           "Control_DB"."Carrousel_Order Table".Task_Data_Available := TRUE;//#System.OrderTable[#Roller_To_Roller_CurrentOrder].OPC_Control.Task_Data_Available; // Send the Task Data Available from WCS 
           "Control_DB"."Carrousel_Order Table".Task_Type := #System.OrderTable[#RTR_P1P2_CurrentOrder].OPC_Control.Task_Type; //  Send the Task Type - Roller to Roller Conveyor = Task Type = 6
           "Control_DB"."Carrousel_Order Table".Task_ID := #System.OrderTable[#RTR_P1P2_CurrentOrder].OPC_Control.Task_ID; // Send the Task ID number;
           "Control_DB"."Carrousel_Order Table".Task_Metadata := #System.OrderTable[#RTR_P1P2_CurrentOrder].OPC_Control.Task_Metadata; // Send the Task Metadata Unique identifier
           "Control_DB"."Carrousel_Order Table".Source_Location := #System.OrderTable[#RTR_P1P2_CurrentOrder].OPC_Control.Source_Location; // Send the Source Location from the Conveyor
           "Control_DB"."Carrousel_Order Table".Destination_Location := #System.OrderTable[#RTR_P1P2_CurrentOrder].OPC_Control.Destination_Location; // Send the Destination Location to the Conveyor;
           #RTR_P1P2_WatchdogStart := true;


       END_IF;

       //RUNNING
       IF (#Cnv_PopUp_1.Running OR #Cnv_PopUp_2.Running) AND #System.Auto_Man THEN
           #System.OrderTable[#RTR_P1P2_CurrentOrder].Status := #RUNNING_STATUS;
       END_IF;

       //Cancel order
       IF #Canceling AND NOT (#Cnv_PopUp_1.Running OR #Cnv_PopUp_2.Running) AND #RTR_P1P2_CurrentOrder <> 0
       THEN
           #System.OrderTable[#RTR_P1P2_CurrentOrder].Status := #CANCELED_STATUS;
           #System.OrderTable[#RTR_P1P2_CurrentOrder].CompleteTime := #CurrentTime;
           #RTR_P1P2_CurrentOrder := 0;

           "Control_DB"."Profiling Station".Start := FALSE;

           "Control_DB"."Carrousel_Order Table".Task_Data_Available := FALSE; // Send the Task Data Available from WCS 
           "Control_DB"."Carrousel_Order Table".Task_Type := 0; //  Send the Task Type - Roller to Roller Conveyor = Task Type = 6
           "Control_DB"."Carrousel_Order Table".Task_ID := 0; // Send the Task ID number;
           "Control_DB"."Carrousel_Order Table".Task_Metadata := ''; // Send the Task Metadata Unique identifier
           "Control_DB"."Carrousel_Order Table".Source_Location := 0; // Send the Source Location from the Conveyor
           "Control_DB"."Carrousel_Order Table".Destination_Location := 0; // Send the Destination Location to the Conveyor;

       END_IF;

       //Error
       IF (#Cnv_PopUp_1.Error OR #Cnv_PopUp_2.Error) THEN
           //#Cnv_Entry.Instruction.Execute := FALSE;
           "Control_DB"."Profiling Station".Start := FALSE;

           "Control_DB"."Carrousel_Order Table".Task_Data_Available := FALSE; // Send the Task Data Available from WCS 
           "Control_DB"."Carrousel_Order Table".Task_Type := 0; //  Send the Task Type - Roller to Roller Conveyor = Task Type = 6
           "Control_DB"."Carrousel_Order Table".Task_ID := 0; // Send the Task ID number;
           "Control_DB"."Carrousel_Order Table".Task_Metadata := ''; // Send the Task Metadata Unique identifier
           "Control_DB"."Carrousel_Order Table".Source_Location := 0; // Send the Source Location from the Conveyor
           "Control_DB"."Carrousel_Order Table".Destination_Location := 0; // Send the Destination Location to the Conveyor;
           #System.OrderTable[#RTR_P1P2_CurrentOrder].ErrorID := (#Cnv_PopUp_1.Cnv_Errors.Error_Word_1
           OR #Cnv_PopUp_2.Cnv_Errors.Error_Word_1)
       ;

       END_IF;

       //MOVEMENT FINALIZED
       #RTR_P1P2DoneRTrig(CLK := "Control_DB".Movement_Completed.RTR_P1TP2);
       IF #RTR_P1P2DoneRTrig.Q THEN
           "Control_DB".Movement_Completed.RTR_P1TP2 := FALSE;
           "Control_DB"."Profiling Station".Start := FALSE;

           "Control_DB"."Carrousel_Order Table".Task_Data_Available := FALSE; // Send the Task Data Available from WCS 
           "Control_DB"."Carrousel_Order Table".Task_Type := 0; //  Send the Task Type - Roller to Roller Conveyor = Task Type = 6
           "Control_DB"."Carrousel_Order Table".Task_ID := 0; // Send the Task ID number;
           "Control_DB"."Carrousel_Order Table".Task_Metadata := ''; // Send the Task Metadata Unique identifier
           "Control_DB"."Carrousel_Order Table".Source_Location := 0; // Send the Source Location from the Conveyor
           "Control_DB"."Carrousel_Order Table".Destination_Location := 0; // Send the Destination Location to the Conveyor;

           #RTR_P1P2_WatchdogStart := FALSE;
           #System.OrderTable[#RTR_P1P2_CurrentOrder].Status := #COMPLETED_STATUS;
           #System.OrderTable[#RTR_P1P2_CurrentOrder].CompleteTime := #CurrentTime;
           #RTR_P1P2_CurrentOrder := 0;
       END_IF;
   END_REGION

   REGION Roller TO Roller - Carousel Conveyors - PP3 PP4
       //Roller conveyors
       IF #System.OrderTable[1].StepNo <> 0
           AND #System.OrderTable[1].Device = #RTR_P3_TO_P4
           AND #System.OrderTable[1].Status = #QUEUED_STATUS
           AND NOT (#Cnv_PopUp_3.Running OR #Cnv_PopUp_4.Running)
           AND NOT #System.Error
           AND NOT #Canceling

       THEN
           #RTR_P3P4_CurrentOrder := 1;
       END_IF;
       IF #System.OrderTable[#RTR_P3P4_CurrentOrder].StepNo <> 0
           AND #System.OrderTable[#RTR_P3P4_CurrentOrder].Device = #RTR_P3_TO_P4
           AND #System.OrderTable[#RTR_P3P4_CurrentOrder].Status = #QUEUED_STATUS
           AND NOT (#Cnv_PopUp_3.Running OR #Cnv_PopUp_4.Running)
           AND NOT #System.Error
           AND NOT #Canceling

       THEN
           //OPC Commands to Move Pallets - Carousel Conveyors
           // WCS => Order Table => OPC Ua Control Table


           "Control_DB"."Carrousel_Order Table".Task_Data_Available := TRUE;//#System.OrderTable[#Roller_To_Roller_CurrentOrder].OPC_Control.Task_Data_Available; // Send the Task Data Available from WCS 
           "Control_DB"."Carrousel_Order Table".Task_Type := #System.OrderTable[#RTR_P3P4_CurrentOrder].OPC_Control.Task_Type; //  Send the Task Type - Roller to Roller Conveyor = Task Type = 6
           "Control_DB"."Carrousel_Order Table".Task_ID := #System.OrderTable[#RTR_P3P4_CurrentOrder].OPC_Control.Task_ID; // Send the Task ID number;
           "Control_DB"."Carrousel_Order Table".Task_Metadata := #System.OrderTable[#RTR_P3P4_CurrentOrder].OPC_Control.Task_Metadata; // Send the Task Metadata Unique identifier
           "Control_DB"."Carrousel_Order Table".Source_Location := #System.OrderTable[#RTR_P3P4_CurrentOrder].OPC_Control.Source_Location; // Send the Source Location from the Conveyor
           "Control_DB"."Carrousel_Order Table".Destination_Location := #System.OrderTable[#RTR_P3P4_CurrentOrder].OPC_Control.Destination_Location; // Send the Destination Location to the Conveyor;
           #RTR_P3P4_WatchdogStart := true;


       END_IF;

       //RUNNING
       IF (#Cnv_PopUp_4.Running OR #Cnv_PopUp_3.Running) AND #System.Auto_Man THEN
           #System.OrderTable[#RTR_P3P4_CurrentOrder].Status := #RUNNING_STATUS;
       END_IF;

       //Cancel order
       IF #Canceling AND NOT (#Cnv_PopUp_4.Running OR #Cnv_PopUp_3.Running) AND #RTR_P3P4_CurrentOrder <> 0
       THEN
           #System.OrderTable[#RTR_P3P4_CurrentOrder].Status := #CANCELED_STATUS;
           #System.OrderTable[#RTR_P3P4_CurrentOrder].CompleteTime := #CurrentTime;
           #RTR_P3P4_CurrentOrder := 0;


           "Control_DB"."Carrousel_Order Table".Task_Data_Available := FALSE; // Send the Task Data Available from WCS 
           "Control_DB"."Carrousel_Order Table".Task_Type := 0; //  Send the Task Type - Roller to Roller Conveyor = Task Type = 6
           "Control_DB"."Carrousel_Order Table".Task_ID := 0; // Send the Task ID number;
           "Control_DB"."Carrousel_Order Table".Task_Metadata := ''; // Send the Task Metadata Unique identifier
           "Control_DB"."Carrousel_Order Table".Source_Location := 0; // Send the Source Location from the Conveyor
           "Control_DB"."Carrousel_Order Table".Destination_Location := 0; // Send the Destination Location to the Conveyor;

       END_IF;

       //Error
       IF (#Cnv_PopUp_4.Error OR #Cnv_PopUp_3.Error) THEN
           //#Cnv_Entry.Instruction.Execute := FALSE;

           "Control_DB"."Carrousel_Order Table".Task_Data_Available := FALSE; // Send the Task Data Available from WCS 
           "Control_DB"."Carrousel_Order Table".Task_Type := 0; //  Send the Task Type - Roller to Roller Conveyor = Task Type = 6
           "Control_DB"."Carrousel_Order Table".Task_ID := 0; // Send the Task ID number;
           "Control_DB"."Carrousel_Order Table".Task_Metadata := ''; // Send the Task Metadata Unique identifier
           "Control_DB"."Carrousel_Order Table".Source_Location := 0; // Send the Source Location from the Conveyor
           "Control_DB"."Carrousel_Order Table".Destination_Location := 0; // Send the Destination Location to the Conveyor;
           #System.OrderTable[#RTR_P3P4_CurrentOrder].ErrorID := (#Cnv_PopUp_3.Cnv_Errors.Error_Word_1
           OR #Cnv_PopUp_4.Cnv_Errors.Error_Word_1)
           ;

       END_IF;

       //MOVEMENT FINALIZED
       #RTR_P3P4DoneRTrig(CLK := "Control_DB".Movement_Completed.RTR_P3TP4);
       IF #RTR_P3P4DoneRTrig.Q THEN
           "Control_DB".Movement_Completed.RTR_P3TP4 := FALSE;

           "Control_DB"."Carrousel_Order Table".Task_Data_Available := FALSE; // Send the Task Data Available from WCS 
           "Control_DB"."Carrousel_Order Table".Task_Type := 0; //  Send the Task Type - Roller to Roller Conveyor = Task Type = 6
           "Control_DB"."Carrousel_Order Table".Task_ID := 0; // Send the Task ID number;
           "Control_DB"."Carrousel_Order Table".Task_Metadata := ''; // Send the Task Metadata Unique identifier
           "Control_DB"."Carrousel_Order Table".Source_Location := 0; // Send the Source Location from the Conveyor
           "Control_DB"."Carrousel_Order Table".Destination_Location := 0; // Send the Destination Location to the Conveyor;

           #RTR_P3P4_WatchdogStart := FALSE;
           #System.OrderTable[#RTR_P3P4_CurrentOrder].Status := #COMPLETED_STATUS;
           #System.OrderTable[#RTR_P3P4_CurrentOrder].CompleteTime := #CurrentTime;
           #RTR_P3P4_CurrentOrder := 0;
       END_IF;
   END_REGION

   REGION Roller TO Roller - Carousel Conveyors - PP4 to outbound
       //Roller conveyors
       IF #System.OrderTable[1].StepNo <> 0
           AND #System.OrderTable[1].Device = #RTR_P4TO
           AND #System.OrderTable[1].Status = #QUEUED_STATUS
           AND NOT (#Cnv_PopUp_4.Running OR #Cnv_Exit.Running)
           AND NOT #System.Error
           AND NOT #Canceling

       THEN
           #RTR_P4TO_CurrentOrder := 1;
       END_IF;
       IF #System.OrderTable[#RTR_P4TO_CurrentOrder].StepNo <> 0
           AND #System.OrderTable[#RTR_P4TO_CurrentOrder].Device = #RTR_P4TO
           AND #System.OrderTable[#RTR_P4TO_CurrentOrder].Status = #QUEUED_STATUS
           AND NOT (#Cnv_PopUp_4.Running OR #Cnv_Exit.Running)
           AND NOT #System.Error
           AND NOT #Canceling

       THEN
           //OPC Commands to Move Pallets - Carousel Conveyors
           // WCS => Order Table => OPC Ua Control Table


           "Control_DB"."Carrousel_Order Table".Task_Data_Available := TRUE;//#System.OrderTable[#Roller_To_Roller_CurrentOrder].OPC_Control.Task_Data_Available; // Send the Task Data Available from WCS 
           "Control_DB"."Carrousel_Order Table".Task_Type := #System.OrderTable[#RTR_P4TO_CurrentOrder].OPC_Control.Task_Type; //  Send the Task Type - Roller to Roller Conveyor = Task Type = 6
           "Control_DB"."Carrousel_Order Table".Task_ID := #System.OrderTable[#RTR_P4TO_CurrentOrder].OPC_Control.Task_ID; // Send the Task ID number;
           "Control_DB"."Carrousel_Order Table".Task_Metadata := #System.OrderTable[#RTR_P4TO_CurrentOrder].OPC_Control.Task_Metadata; // Send the Task Metadata Unique identifier
           "Control_DB"."Carrousel_Order Table".Source_Location := #System.OrderTable[#RTR_P4TO_CurrentOrder].OPC_Control.Source_Location; // Send the Source Location from the Conveyor
           "Control_DB"."Carrousel_Order Table".Destination_Location := #System.OrderTable[#RTR_P4TO_CurrentOrder].OPC_Control.Destination_Location; // Send the Destination Location to the Conveyor;
           #RTR_P4TO_WatchdogStart := true;


       END_IF;

       //RUNNING
       IF (#Cnv_PopUp_4.Running OR #Cnv_Exit.Running) AND #System.Auto_Man THEN
           #System.OrderTable[#RTR_P4TO_CurrentOrder].Status := #RUNNING_STATUS;
       END_IF;

       //Cancel order
       IF #Canceling AND NOT (#Cnv_PopUp_4.Running OR #Cnv_Exit.Running) AND #RTR_P4TO_CurrentOrder <> 0
       THEN
           #System.OrderTable[#RTR_P4TO_CurrentOrder].Status := #CANCELED_STATUS;
           #System.OrderTable[#RTR_P4TO_CurrentOrder].CompleteTime := #CurrentTime;
           #RTR_P4TO_CurrentOrder := 0;


           "Control_DB"."Carrousel_Order Table".Task_Data_Available := FALSE; // Send the Task Data Available from WCS 
           "Control_DB"."Carrousel_Order Table".Task_Type := 0; //  Send the Task Type - Roller to Roller Conveyor = Task Type = 6
           "Control_DB"."Carrousel_Order Table".Task_ID := 0; // Send the Task ID number;
           "Control_DB"."Carrousel_Order Table".Task_Metadata := ''; // Send the Task Metadata Unique identifier
           "Control_DB"."Carrousel_Order Table".Source_Location := 0; // Send the Source Location from the Conveyor
           "Control_DB"."Carrousel_Order Table".Destination_Location := 0; // Send the Destination Location to the Conveyor;

       END_IF;

       //Error
       IF (#Cnv_PopUp_4.Error OR #Cnv_Exit.Error) THEN
           //#Cnv_Entry.Instruction.Execute := FALSE;

           "Control_DB"."Carrousel_Order Table".Task_Data_Available := FALSE; // Send the Task Data Available from WCS 
           "Control_DB"."Carrousel_Order Table".Task_Type := 0; //  Send the Task Type - Roller to Roller Conveyor = Task Type = 6
           "Control_DB"."Carrousel_Order Table".Task_ID := 0; // Send the Task ID number;
           "Control_DB"."Carrousel_Order Table".Task_Metadata := ''; // Send the Task Metadata Unique identifier
           "Control_DB"."Carrousel_Order Table".Source_Location := 0; // Send the Source Location from the Conveyor
           "Control_DB"."Carrousel_Order Table".Destination_Location := 0; // Send the Destination Location to the Conveyor;
           #System.OrderTable[#RTR_P3P4_CurrentOrder].ErrorID := (#Cnv_PopUp_3.Cnv_Errors.Error_Word_1
           OR #Cnv_PopUp_4.Cnv_Errors.Error_Word_1)
           ;

       END_IF;

       //MOVEMENT FINALIZED
       #RTR_P4TODoneRTrig(CLK := "Control_DB".Movement_Completed.RTR_P4TO);
       IF #RTR_P4TODoneRTrig.Q THEN
           "Control_DB".Movement_Completed.RTR_P4TO := FALSE;

           "Control_DB"."Carrousel_Order Table".Task_Data_Available := FALSE; // Send the Task Data Available from WCS 
           "Control_DB"."Carrousel_Order Table".Task_Type := 0; //  Send the Task Type - Roller to Roller Conveyor = Task Type = 6
           "Control_DB"."Carrousel_Order Table".Task_ID := 0; // Send the Task ID number;
           "Control_DB"."Carrousel_Order Table".Task_Metadata := ''; // Send the Task Metadata Unique identifier
           "Control_DB"."Carrousel_Order Table".Source_Location := 0; // Send the Source Location from the Conveyor
           "Control_DB"."Carrousel_Order Table".Destination_Location := 0; // Send the Destination Location to the Conveyor;

           #RTR_P4TO_WatchdogStart := FALSE;
           #System.OrderTable[#RTR_P4TO_CurrentOrder].Status := #COMPLETED_STATUS;
           #System.OrderTable[#RTR_P4TO_CurrentOrder].CompleteTime := #CurrentTime;
           #RTR_P4TO_CurrentOrder := 0;
       END_IF;
   END_REGION




   REGION Chain to Chain - Carousel Conveyors - Pop 2 to Pop 3
       IF #System.OrderTable[1].StepNo <> 0
           AND #System.OrderTable[1].Device = #CHAIN_TO_CHAIN_DEVICE
           AND #System.OrderTable[1].Status = #QUEUED_STATUS
           AND NOT (#Cnv_PopUp_2.Running OR #Cnv_PopUp_3.Running)
           AND NOT #System.Error
           AND NOT #Canceling
           //AND #System.OrderTable[#Chain_To_Chain_CurrentOrder].Status <> #RUNNING_STATUS

       THEN
           #Chain_To_Chain_CurrentOrder := 1;
       END_IF;
       IF #System.OrderTable[#Chain_To_Chain_CurrentOrder].StepNo <> 0
           AND #System.OrderTable[#Chain_To_Chain_CurrentOrder].Device = #CHAIN_TO_CHAIN_DEVICE
           AND #System.OrderTable[#Chain_To_Chain_CurrentOrder].Status = #QUEUED_STATUS
           AND NOT (#Cnv_PopUp_2.Running OR #Cnv_PopUp_3.Running)
           AND NOT #System.Error
           AND NOT #Canceling
          // AND #System.OrderTable[#Chain_To_Chain_CurrentOrder].Status <> #RUNNING_STATUS
       THEN
           //OPC Commands to Move Pallets - Carousel Conveyors
           // WCS => Order Table => OPC Ua Control Table

           "Control_DB"."Carrousel_Order Table".Task_Data_Available := TRUE;//#System.OrderTable[#Chain_To_Chain_CurrentOrder].OPC_Control.Task_Data_Available; // Send the Task Data Available from WCS 
           "Control_DB"."Carrousel_Order Table".Task_Type := #System.OrderTable[#Chain_To_Chain_CurrentOrder].OPC_Control.Task_Type; //  Send the Task Type - Chain to Chain Conveyor = Task Type = 7
           "Control_DB"."Carrousel_Order Table".Task_ID := #System.OrderTable[#Chain_To_Chain_CurrentOrder].OPC_Control.Task_ID; // Send the Task ID number;
           "Control_DB"."Carrousel_Order Table".Task_Metadata := #System.OrderTable[#Chain_To_Chain_CurrentOrder].OPC_Control.Task_Metadata; // Send the Task Metadata Unique identifier
           "Control_DB"."Carrousel_Order Table".Source_Location := #System.OrderTable[#Chain_To_Chain_CurrentOrder].OPC_Control.Source_Location; // Send the Source Location from the Conveyor
           "Control_DB"."Carrousel_Order Table".Destination_Location := #System.OrderTable[#Chain_To_Chain_CurrentOrder].OPC_Control.Destination_Location; // Send the Destination Location to the Conveyor;
           #Chain_To_Chain_WatchdogStart := true;


       END_IF;

       //RUNNING
       IF (#Cnv_PopUp_2.Running OR #Cnv_PopUp_3.Running)AND #System.Auto_Man THEN
           //#Cnv_Entry.Instruction.Execute := FALSE;
           #System.OrderTable[#Chain_To_Chain_CurrentOrder].Status := #RUNNING_STATUS;
       END_IF;

       //Cancel order
       IF #Canceling AND NOT (#Cnv_PopUp_2.Running OR #Cnv_PopUp_3.Running) AND #Chain_To_Chain_CurrentOrder <> 0 THEN


           "Control_DB"."Carrousel_Order Table".Task_Data_Available := FALSE;//#System.OrderTable[#Chain_To_Chain_CurrentOrder].OPC_Control.Task_Data_Available; // Send the Task Data Available from WCS 
           "Control_DB"."Carrousel_Order Table".Task_Type := 0; //  Send the Task Type - Chain to Chain Conveyor = Task Type = 7
           "Control_DB"."Carrousel_Order Table".Task_ID := 0; // Send the Task ID number;
           "Control_DB"."Carrousel_Order Table".Task_Metadata := ''; // Send the Task Metadata Unique identifier
           "Control_DB"."Carrousel_Order Table".Source_Location := 0; // Send the Source Location from the Conveyor
           "Control_DB"."Carrousel_Order Table".Destination_Location := 0; // Send the Destination Location to the Conveyor;

           #System.OrderTable[#Chain_To_Chain_CurrentOrder].Status := #CANCELED_STATUS;
           #System.OrderTable[#Chain_To_Chain_CurrentOrder].CompleteTime := #CurrentTime;
           #Chain_To_Chain_CurrentOrder := 0;
           //#Cnv_Entry.Instruction.Execute := FALSE;
       END_IF;

       //Error
       IF (#Cnv_PopUp_2.Error OR #Cnv_PopUp_3.Error) THEN
           //#Cnv_Entry.Instruction.Execute := FALSE;
           //
           "Control_DB"."Carrousel_Order Table".Task_Data_Available := FALSE;//#System.OrderTable[#Chain_To_Chain_CurrentOrder].OPC_Control.Task_Data_Available; // Send the Task Data Available from WCS 
           "Control_DB"."Carrousel_Order Table".Task_Type := 0; //  Send the Task Type - Chain to Chain Conveyor = Task Type = 7
           "Control_DB"."Carrousel_Order Table".Task_ID := 0; // Send the Task ID number;
           "Control_DB"."Carrousel_Order Table".Task_Metadata := ''; // Send the Task Metadata Unique identifier
           "Control_DB"."Carrousel_Order Table".Source_Location := 0; // Send the Source Location from the Conveyor
           "Control_DB"."Carrousel_Order Table".Destination_Location := 0; // Send the Destination Location to the Conveyor;

           #System.OrderTable[#Chain_To_Chain_CurrentOrder].ErrorID := (#Cnv_PopUp_2.Cnv_Errors.Error_Word_1
                                                                        OR #Cnv_PopUp_3.Cnv_Errors.Error_Word_1);

       END_IF;

       //MOVEMENT FINALIZED
       #Chain_To_ChainDoneRTrig(CLK := "Control_DB".Movement_Completed.RTR_P2TP3);
       IF #Chain_To_ChainDoneRTrig.Q THEN
           "Control_DB".Movement_Completed.RTR_P2TP3 := FALSE;
           "Control_DB"."Carrousel_Order Table".Task_Data_Available := FALSE;//#System.OrderTable[#Chain_To_Chain_CurrentOrder].OPC_Control.Task_Data_Available; // Send the Task Data Available from WCS 
           "Control_DB"."Carrousel_Order Table".Task_Type := 0; //  Send the Task Type - Chain to Chain Conveyor = Task Type = 7
           "Control_DB"."Carrousel_Order Table".Task_ID := 0; // Send the Task ID number;
           "Control_DB"."Carrousel_Order Table".Task_Metadata := ''; // Send the Task Metadata Unique identifier
           "Control_DB"."Carrousel_Order Table".Source_Location := 0; // Send the Source Location from the Conveyor
           "Control_DB"."Carrousel_Order Table".Destination_Location := 0; // Send the Destination Location to the Conveyor;


           #Chain_To_Chain_WatchdogStart := FALSE;
           #System.OrderTable[#Chain_To_Chain_CurrentOrder].Status := #COMPLETED_STATUS;
           #System.OrderTable[#Chain_To_Chain_CurrentOrder].CompleteTime := #CurrentTime;
           #Chain_To_Chain_CurrentOrder := 0;
       END_IF;
   END_REGION

   REGION Pop4 to Pick Station - Carousel Conveyors - Pop 4 to Pick Station
       IF #System.OrderTable[1].StepNo <> 0
           AND #System.OrderTable[1].Device = #POP4_TO_PICK_DEVICE
           AND #System.OrderTable[1].Status = #QUEUED_STATUS
          // AND NOT "Control_DB".Pick_Station.Running
           AND NOT #System.Error
           AND NOT #Canceling
           AND #System.OrderTable[1].Status <> #RUNNING_STATUS
           //AND #System.OrderTable[#PickSt_To_Pop1_CurrentOrder].Status <> #RUNNING_STATUS

       THEN
           #Pop4_To_PickSt_CurrentOrder := 1;
       END_IF;
       IF #System.OrderTable[#Pop4_To_PickSt_CurrentOrder].StepNo <> 0
           AND #System.OrderTable[#Pop4_To_PickSt_CurrentOrder].Device = #POP4_TO_PICK_DEVICE
           AND #System.OrderTable[#Pop4_To_PickSt_CurrentOrder].Status = #QUEUED_STATUS
           // AND NOT "Control_DB".Pick_Station.Running
           AND NOT #System.Error
           AND NOT #Canceling
           AND #System.OrderTable[#Pop4_To_PickSt_CurrentOrder].Status <> #RUNNING_STATUS
           //AND #System.OrderTable[#PickSt_To_Pop1_CurrentOrder].Status <> #RUNNING_STATUS
       THEN
           //OPC Commands to Move Pallets - Carousel Conveyors
           // WCS => Order Table => OPC Ua Control Table

           "Control_DB"."Carrousel_Order Table".Task_Data_Available := TRUE;//#System.OrderTable[#Pop4_To_PickSt_CurrentOrder].OPC_Control.Task_Data_Available; // Send the Task Data Available from WCS 
           "Control_DB"."Carrousel_Order Table".Task_Type := #System.OrderTable[#Pop4_To_PickSt_CurrentOrder].OPC_Control.Task_Type; //  Send the Task Type - Pop4 to Pick Station Conveyor = Task Type = 8
           "Control_DB"."Carrousel_Order Table".Task_ID := #System.OrderTable[#Pop4_To_PickSt_CurrentOrder].OPC_Control.Task_ID; // Send the Task ID number;
           "Control_DB"."Carrousel_Order Table".Task_Metadata := #System.OrderTable[#Pop4_To_PickSt_CurrentOrder].OPC_Control.Task_Metadata; // Send the Task Metadata Unique identifier
           "Control_DB"."Carrousel_Order Table".Source_Location := #System.OrderTable[#Pop4_To_PickSt_CurrentOrder].OPC_Control.Source_Location; // Send the Source Location from the Conveyor
           "Control_DB"."Carrousel_Order Table".Destination_Location := #System.OrderTable[#Pop4_To_PickSt_CurrentOrder].OPC_Control.Destination_Location; // Send the Destination Location to the Conveyor;
           #Pop4_To_PickWatchdogStart := TRUE;



       END_IF;

       //RUNNING
       IF "Control_DB".Pick_Station.Running AND #System.Auto_Man THEN
           //#Cnv_Entry.Instruction.Execute := FALSE;
           #System.OrderTable[#Pop4_To_PickSt_CurrentOrder].Status := #RUNNING_STATUS;
       END_IF;

       //Cancel order
       IF #Canceling AND NOT "Control_DB".Pick_Station.Running AND #Pop4_To_PickSt_CurrentOrder <> 0 THEN
           #System.OrderTable[#Pop4_To_PickSt_CurrentOrder].Status := #CANCELED_STATUS;
           #System.OrderTable[#Pop4_To_PickSt_CurrentOrder].CompleteTime := #CurrentTime;
           #Pop4_To_PickSt_CurrentOrder := 0;

           "Control_DB"."Carrousel_Order Table".Task_Data_Available := FALSE;//#System.OrderTable[#Chain_To_Chain_CurrentOrder].OPC_Control.Task_Data_Available; // Send the Task Data Available from WCS 
           "Control_DB"."Carrousel_Order Table".Task_Type := 0; //  Send the Task Type - Chain to Chain Conveyor = Task Type = 7
           "Control_DB"."Carrousel_Order Table".Task_ID := 0; // Send the Task ID number;
           "Control_DB"."Carrousel_Order Table".Task_Metadata := ''; // Send the Task Metadata Unique identifier
           "Control_DB"."Carrousel_Order Table".Source_Location := 0; // Send the Source Location from the Conveyor
           "Control_DB"."Carrousel_Order Table".Destination_Location := 0; // Send the Destination Location to the Conveyor;

           //#Cnv_Entry.Instruction.Execute := FALSE;
       END_IF;

       //Error
       IF "Control_DB".Pick_Station.Error THEN
           //#Cnv_Entry.Instruction.Execute := FALSE;
           "Control_DB"."Carrousel_Order Table".Task_Data_Available := FALSE;//#System.OrderTable[#Chain_To_Chain_CurrentOrder].OPC_Control.Task_Data_Available; // Send the Task Data Available from WCS 
           "Control_DB"."Carrousel_Order Table".Task_Type := 0; //  Send the Task Type - Chain to Chain Conveyor = Task Type = 7
           "Control_DB"."Carrousel_Order Table".Task_ID := 0; // Send the Task ID number;
           "Control_DB"."Carrousel_Order Table".Task_Metadata := ''; // Send the Task Metadata Unique identifier
           "Control_DB"."Carrousel_Order Table".Source_Location := 0; // Send the Source Location from the Conveyor
           "Control_DB"."Carrousel_Order Table".Destination_Location := 0; // Send the Destination Location to the Conveyor;
           #System.OrderTable[#Pop4_To_PickSt_CurrentOrder].ErrorID := "Control_DB".Pick_Station.Cnv_Errors.Error_Word_1;

       END_IF;

       //MOVEMENT FINALIZED
       #Pop4_To_PickSt_DoneRTrig(CLK := "Control_DB".Movement_Completed.Pop4_To_Pick);
       IF #Pop4_To_PickSt_DoneRTrig.Q THEN
           "Control_DB".Movement_Completed.Pop4_To_Pick := FALSE;
           #Pop4_To_PickWatchdogStart := FALSE;

           "Control_DB"."Carrousel_Order Table".Task_Data_Available := FALSE;//#System.OrderTable[#Chain_To_Chain_CurrentOrder].OPC_Control.Task_Data_Available; // Send the Task Data Available from WCS 
           "Control_DB"."Carrousel_Order Table".Task_Type := 0; //  Send the Task Type - Chain to Chain Conveyor = Task Type = 7
           "Control_DB"."Carrousel_Order Table".Task_ID := 0; // Send the Task ID number;
           "Control_DB"."Carrousel_Order Table".Task_Metadata := ''; // Send the Task Metadata Unique identifier
           "Control_DB"."Carrousel_Order Table".Source_Location := 0; // Send the Source Location from the Conveyor
           "Control_DB"."Carrousel_Order Table".Destination_Location := 0; // Send the Destination Location to the Conveyor;

           #System.OrderTable[#Pop4_To_PickSt_CurrentOrder].Status := #COMPLETED_STATUS;
           #System.OrderTable[#Pop4_To_PickSt_CurrentOrder].CompleteTime := #CurrentTime;
           #Pop4_To_PickSt_CurrentOrder := 0;
       END_IF;
   END_REGION

   REGION Pick Station to Pop1 - Carousel Conveyors - Pick Station To Pop 1 
       IF #System.OrderTable[1].StepNo <> 0
           AND #System.OrderTable[1].Device = #PICK_TO_POP1_DEVICE
           AND #System.OrderTable[1].Status = #QUEUED_STATUS
           AND NOT (#Cnv_PopUp_1.Running)
           AND NOT #System.Error
           AND NOT #Canceling
           //AND #System.OrderTable[#Roller_To_Roller_CurrentOrder].Status <> #RUNNING_STATUS
           //AND #System.OrderTable[#Pop4_To_PickSt_CurrentOrder].Status <> #RUNNING_STATUS
       THEN
           #PickSt_To_Pop1_CurrentOrder := 1;
       END_IF;
       IF #System.OrderTable[#PickSt_To_Pop1_CurrentOrder].StepNo <> 0
           AND #System.OrderTable[#PickSt_To_Pop1_CurrentOrder].Device = #PICK_TO_POP1_DEVICE
           AND #System.OrderTable[#PickSt_To_Pop1_CurrentOrder].Status = #QUEUED_STATUS
           AND NOT (#Cnv_PopUp_1.Running)
           AND NOT #System.Error
           AND NOT #Canceling
           //AND #System.OrderTable[#Roller_To_Roller_CurrentOrder].Status <> #RUNNING_STATUS
           //AND #System.OrderTable[#Pop4_To_PickSt_CurrentOrder].Status <> #RUNNING_STATUS
       THEN
           //OPC Commands to Move Pallets - Carousel Conveyors
           // WCS => Order Table => OPC Ua Control Table

           "Control_DB"."Carrousel_Order Table".Task_Data_Available := TRUE;//#System.OrderTable[#PickSt_To_Pop1_CurrentOrder].OPC_Control.Task_Data_Available; // Send the Task Data Available from WCS 
           "Control_DB"."Carrousel_Order Table".Task_Type := #System.OrderTable[#PickSt_To_Pop1_CurrentOrder].OPC_Control.Task_Type; //  Send the Task Type - Roller to Roller Conveyor = Task Type = 6
           "Control_DB"."Carrousel_Order Table".Task_ID := #System.OrderTable[#PickSt_To_Pop1_CurrentOrder].OPC_Control.Task_ID; // Send the Task ID number;
           "Control_DB"."Carrousel_Order Table".Task_Metadata := #System.OrderTable[#PickSt_To_Pop1_CurrentOrder].OPC_Control.Task_Metadata; // Send the Task Metadata Unique identifier
           "Control_DB"."Carrousel_Order Table".Source_Location := #System.OrderTable[#PickSt_To_Pop1_CurrentOrder].OPC_Control.Source_Location; // Send the Source Location from the Conveyor
           "Control_DB"."Carrousel_Order Table".Destination_Location := #System.OrderTable[#PickSt_To_Pop1_CurrentOrder].OPC_Control.Destination_Location; // Send the Destination Location to the Conveyor;
           #PickSt_To_Pop1WatchdogStart := true;


       END_IF;

       //RUNNING
       IF (#Cnv_PopUp_1.Running) AND #System.Auto_Man THEN
           //#Cnv_Entry.Instruction.Execute := FALSE;
           #System.OrderTable[#PickSt_To_Pop1_CurrentOrder].Status := #RUNNING_STATUS;
       END_IF;

       //Cancel order
       IF #Canceling AND NOT (#Cnv_PopUp_1.Running) AND #PickSt_To_Pop1_CurrentOrder <> 0 THEN
           #System.OrderTable[#PickSt_To_Pop1_CurrentOrder].Status := #CANCELED_STATUS;
           #System.OrderTable[#PickSt_To_Pop1_CurrentOrder].CompleteTime := #CurrentTime;
           #PickSt_To_Pop1_CurrentOrder := 0;
           "Control_DB"."Carrousel_Order Table".Task_Data_Available := FALSE;//#System.OrderTable[#Chain_To_Chain_CurrentOrder].OPC_Control.Task_Data_Available; // Send the Task Data Available from WCS 
           "Control_DB"."Carrousel_Order Table".Task_Type := 0; //  Send the Task Type - Chain to Chain Conveyor = Task Type = 7
           "Control_DB"."Carrousel_Order Table".Task_ID := 0; // Send the Task ID number;
           "Control_DB"."Carrousel_Order Table".Task_Metadata := ''; // Send the Task Metadata Unique identifier
           "Control_DB"."Carrousel_Order Table".Source_Location := 0; // Send the Source Location from the Conveyor
           "Control_DB"."Carrousel_Order Table".Destination_Location := 0; // Send the Destination Location to the Conveyor;
           //#Cnv_Entry.Instruction.Execute := FALSE;
       END_IF;

       //Error
       IF (#Cnv_PopUp_2.Error OR #Cnv_PopUp_3.Error) THEN
           //#Cnv_Entry.Instruction.Execute := FALSE;
           "Control_DB"."Carrousel_Order Table".Task_Data_Available := FALSE;//#System.OrderTable[#Chain_To_Chain_CurrentOrder].OPC_Control.Task_Data_Available; // Send the Task Data Available from WCS 
           "Control_DB"."Carrousel_Order Table".Task_Type := 0; //  Send the Task Type - Chain to Chain Conveyor = Task Type = 7
           "Control_DB"."Carrousel_Order Table".Task_ID := 0; // Send the Task ID number;
           "Control_DB"."Carrousel_Order Table".Task_Metadata := ''; // Send the Task Metadata Unique identifier
           "Control_DB"."Carrousel_Order Table".Source_Location := 0; // Send the Source Location from the Conveyor
           "Control_DB"."Carrousel_Order Table".Destination_Location := 0; // Send the Destination Location to the Conveyor;
           #System.OrderTable[#PickSt_To_Pop1_CurrentOrder].ErrorID := (#Cnv_PopUp_2.Cnv_Errors.Error_Word_1
           OR #Cnv_PopUp_3.Cnv_Errors.Error_Word_1);

       END_IF;

       //MOVEMENT FINALIZED
       #PickSt_To_Pop1_DoneRTrig(CLK := "Control_DB".Movement_Completed.Pick_To_Pop1);
       IF #PickSt_To_Pop1_DoneRTrig.Q THEN
           "Control_DB".Movement_Completed.Pick_To_Pop1 := FALSE;
           "Control_DB"."Carrousel_Order Table".Task_Data_Available := FALSE;//#System.OrderTable[#Chain_To_Chain_CurrentOrder].OPC_Control.Task_Data_Available; // Send the Task Data Available from WCS 
           "Control_DB"."Carrousel_Order Table".Task_Type := 0; //  Send the Task Type - Chain to Chain Conveyor = Task Type = 7
           "Control_DB"."Carrousel_Order Table".Task_ID := 0; // Send the Task ID number;
           "Control_DB"."Carrousel_Order Table".Task_Metadata := ''; // Send the Task Metadata Unique identifier
           "Control_DB"."Carrousel_Order Table".Source_Location := 0; // Send the Source Location from the Conveyor
           "Control_DB"."Carrousel_Order Table".Destination_Location := 0; // Send the Destination Location to the Conveyor;

           #PickSt_To_Pop1WatchdogStart := FALSE;
           #System.OrderTable[#PickSt_To_Pop1_CurrentOrder].Status := #COMPLETED_STATUS;
           #System.OrderTable[#PickSt_To_Pop1_CurrentOrder].CompleteTime := #CurrentTime;
           #PickSt_To_Pop1_CurrentOrder := 0;
       END_IF;
   END_REGION

   REGION Weigh Station - Carousel Conveyors 
       IF #System.OrderTable[1].StepNo <> 0
           AND #System.OrderTable[1].Device = #WEIGH_STATION_DEVICE
           AND #System.OrderTable[1].Status = #QUEUED_STATUS
           AND NOT ("Control_DB"."Weighing Station".Running)
           AND NOT #System.Error
           AND NOT #Canceling
       THEN
           #WeighingStation_CurrentOrder := 1;
       END_IF;
       IF #System.OrderTable[#WeighingStation_CurrentOrder].StepNo <> 0
           AND #System.OrderTable[#WeighingStation_CurrentOrder].Device = #WEIGH_STATION_DEVICE
           AND #System.OrderTable[#WeighingStation_CurrentOrder].Status = #QUEUED_STATUS
           AND NOT ("Control_DB"."Weighing Station".Running)
           AND NOT #System.Error
           AND NOT #Canceling
       THEN
           //OPC Commands to Move Pallets - Carousel Conveyors
           // WCS => Order Table => OPC Ua Control Table


           "Control_DB"."Carrousel_Order Table".Task_Data_Available := TRUE;//#System.OrderTable[#WeighingStation_CurrentOrder].OPC_Control.Task_Data_Available; // Send the Task Data Available from WCS 
           "Control_DB"."Carrousel_Order Table".Task_Type := #System.OrderTable[#WeighingStation_CurrentOrder].OPC_Control.Task_Type; //  Send the Task Type - Start Weigh Station = Task Type = 10
           "Control_DB"."Carrousel_Order Table".Task_ID := #System.OrderTable[#WeighingStation_CurrentOrder].OPC_Control.Task_ID; // Send the Task ID number;
           "Control_DB"."Carrousel_Order Table".Task_Metadata := #System.OrderTable[#WeighingStation_CurrentOrder].OPC_Control.Task_Metadata; // Send the Task Metadata Unique identifier
           #WeighingStation_WatchdogStart := true;


       END_IF;

       //RUNNING
       IF ("Control_DB"."Weighing Station".Running) AND #System.Auto_Man
           (*AND NOT "Control_DB".Movement_Completed.WeighingStation*) THEN
           //#Cnv_Entry.Instruction.Execute := FALSE;
           #System.OrderTable[#WeighingStation_CurrentOrder].Status := #RUNNING_STATUS;
           "Control_DB"."Carrousel_Order Table".Task_Data_Available := FALSE;
       END_IF;

       //Cancel order
       IF #Canceling AND NOT ("Control_DB"."Weighing Station".Running) AND #WeighingStation_CurrentOrder <> 0 THEN
           #System.OrderTable[#WeighingStation_CurrentOrder].Status := #CANCELED_STATUS;
           #System.OrderTable[#WeighingStation_CurrentOrder].CompleteTime := #CurrentTime;
           #WeighingStation_CurrentOrder := 0;
           //#Cnv_Entry.Instruction.Execute := FALSE;
           "Control_DB"."Carrousel_Order Table".Task_Data_Available := FALSE;//#System.OrderTable[#WeighingStation_CurrentOrder].OPC_Control.Task_Data_Available; // Send the Task Data Available from WCS 
           "Control_DB"."Carrousel_Order Table".Task_Type := 0; //  Send the Task Type - Start Weigh Station = Task Type = 10
           "Control_DB"."Carrousel_Order Table".Task_ID := 0; // Send the Task ID number;
           "Control_DB"."Carrousel_Order Table".Task_Metadata := ''; // Send the Task Metadata Unique identifier
       END_IF;
     (*  
       //Error
       IF (#WeighingStation. OR #Cnv_PopUp_3.Error) THEN
           //#Cnv_Entry.Instruction.Execute := FALSE;

           #System.OrderTable[#WeighingStation_CurrentOrder].ErrorID := (#Cnv_PopUp_2.Cnv_Errors.Error_Word_1
         OR #Cnv_PopUp_3.Cnv_Errors.Error_Word_1);

       END_IF;
      *) 
       //MOVEMENT FINALIZED
       #WeighingStationDoneRTrig(CLK := "Control_DB".Movement_Completed.WeighingStation);
       IF #WeighingStationDoneRTrig.Q THEN
           "Control_DB".Movement_Completed.WeighingStation := FALSE;
           #WeighingStation_WatchdogStart := FALSE;
           #System.OrderTable[#WeighingStation_CurrentOrder].Status := #COMPLETED_STATUS;
           #System.OrderTable[#WeighingStation_CurrentOrder].CompleteTime := #CurrentTime;
           #WeighingStation_CurrentOrder := 0;

           "Control_DB"."Carrousel_Order Table".Task_Data_Available := FALSE;//#System.OrderTable[#WeighingStation_CurrentOrder].OPC_Control.Task_Data_Available; // Send the Task Data Available from WCS 
           "Control_DB"."Carrousel_Order Table".Task_Type := 0; //  Send the Task Type - Start Weigh Station = Task Type = 10
           "Control_DB"."Carrousel_Order Table".Task_ID := 0; // Send the Task ID number;
           "Control_DB"."Carrousel_Order Table".Task_Metadata := ''; // Send the Task Metadata Unique identifier
       END_IF;
   END_REGION
   (*
   REGION Profile Station - Carousel Conveyors 
       IF #System.OrderTable[1].StepNo <> 0
           AND #System.OrderTable[1].Device = #PROFILE_STATION_DEVICE
           AND #System.OrderTable[1].Status = #QUEUED_STATUS
           AND NOT ("Control_DB"."Profiling Station".Running)
           AND NOT #System.Error
           AND NOT #Canceling
       THEN
           #ProfileStation_CurrentOrder := 1;
       END_IF;
       IF #System.OrderTable[#ProfileStation_CurrentOrder].StepNo <> 0
           AND #System.OrderTable[#ProfileStation_CurrentOrder].Device = #PROFILE_STATION_DEVICE
           AND #System.OrderTable[#ProfileStation_CurrentOrder].Status = #QUEUED_STATUS
           AND NOT ("Control_DB"."Profiling Station".Running)
           AND NOT #System.Error
           AND NOT #Canceling
       THEN
           //OPC Commands to Move Pallets - Carousel Conveyors
           // WCS => Order Table => OPC Ua Control Table

           "Control_DB"."Carrousel_Order Table".Task_Data_Available := TRUE;//#System.OrderTable[#ProfileStation_CurrentOrder].OPC_Control.Task_Data_Available; // Send the Task Data Available from WCS 
           "Control_DB"."Carrousel_Order Table".Task_Type := #System.OrderTable[#ProfileStation_CurrentOrder].OPC_Control.Task_Type; //  Send the Task Type - Start Weigh Station = Task Type = 10
           "Control_DB"."Carrousel_Order Table".Task_ID := #System.OrderTable[#ProfileStation_CurrentOrder].OPC_Control.Task_ID; // Send the Task ID number;
           "Control_DB"."Carrousel_Order Table".Task_Metadata := #System.OrderTable[#ProfileStation_CurrentOrder].OPC_Control.Task_Metadata; // Send the Task Metadata Unique identifier
           #ProfileStation_WatchdogStart := true;


       END_IF;

       //RUNNING
       IF ("Control_DB"."Profiling Station".Running) AND #System.Auto_Man THEN
           //#Cnv_Entry.Instruction.Execute := FALSE;
           #System.OrderTable[#ProfileStation_CurrentOrder].Status := #RUNNING_STATUS;

           "Control_DB"."Carrousel_Order Table".Task_Data_Available := FALSE;//#System.OrderTable[#ProfileStation_CurrentOrder].OPC_Control.Task_Data_Available; // Send the Task Data Available from WCS 
           "Control_DB"."Carrousel_Order Table".Task_Type := 0; //  Send the Task Type - Start Weigh Station = Task Type = 10
           "Control_DB"."Carrousel_Order Table".Task_ID := 0; // Send the Task ID number;
           "Control_DB"."Carrousel_Order Table".Task_Metadata := ''; // Send the Task Metadata Unique identifier
           #ProfileStation_WatchdogStart := true;
       END_IF;

       //Cancel order
       IF #Canceling AND NOT ("Control_DB"."Profiling Station".Running) AND #ProfileStation_CurrentOrder <> 0 THEN
           #System.OrderTable[#ProfileStation_CurrentOrder].Status := #CANCELED_STATUS;
           #System.OrderTable[#ProfileStation_CurrentOrder].CompleteTime := #CurrentTime;
           #ProfileStation_CurrentOrder := 0;
           "Control_DB"."Carrousel_Order Table".Task_Data_Available := FALSE;//#System.OrderTable[#ProfileStation_CurrentOrder].OPC_Control.Task_Data_Available; // Send the Task Data Available from WCS 
           "Control_DB"."Carrousel_Order Table".Task_Type := 0; //  Send the Task Type - Start Weigh Station = Task Type = 10
           "Control_DB"."Carrousel_Order Table".Task_ID := 0; // Send the Task ID number;
           "Control_DB"."Carrousel_Order Table".Task_Metadata := ''; // Send the Task Metadata Unique identifier
           //#Cnv_Entry.Instruction.Execute := FALSE;
       END_IF;
       (*  
         //Error
         IF (#WeighingStation. OR #Cnv_PopUp_3.Error) THEN
             //#Cnv_Entry.Instruction.Execute := FALSE;

             #System.OrderTable[#WeighingStation_CurrentOrder].ErrorID := (#Cnv_PopUp_2.Cnv_Errors.Error_Word_1
           OR #Cnv_PopUp_3.Cnv_Errors.Error_Word_1);

         END_IF;
        *)
        //MOVEMENT FINALIZED
       #ProfileStationDoneRTrig(CLK := "Control_DB"."Profiling Station".Done);
       IF #ProfileStationDoneRTrig.Q THEN
            #ProfileStation_WatchdogStart := FALSE;
            #System.OrderTable[#ProfileStation_CurrentOrder].Status := #COMPLETED_STATUS;
            #System.OrderTable[#ProfileStation_CurrentOrder].CompleteTime := #CurrentTime;
            #ProfileStation_CurrentOrder := 0;
            "Control_DB"."Carrousel_Order Table".Task_Data_Available := FALSE;//#System.OrderTable[#ProfileStation_CurrentOrder].OPC_Control.Task_Data_Available; // Send the Task Data Available from WCS 
            "Control_DB"."Carrousel_Order Table".Task_Type := 0; //  Send the Task Type - Start Weigh Station = Task Type = 10
            "Control_DB"."Carrousel_Order Table".Task_ID := 0; // Send the Task ID number;
            "Control_DB"."Carrousel_Order Table".Task_Metadata := ''; // Send the Task Metadata Unique identifier
        END_IF;
    END_REGION
   *)
   REGION Max Running Order Number
       #MaxRunningOrderNo := MAX(IN1 := #Roller_To_Roller_CurrentOrder, IN2 := #Chain_To_Chain_CurrentOrder,
                                 IN3 := #Pop4_To_PickSt_CurrentOrder, IN4 := #PickSt_To_Pop1_CurrentOrder,
                                 IN5 := #WeighingStation_CurrentOrder, IN6 := #ProfileStation_CurrentOrder);
   END_REGION

   REGION Pause Orders
       #ErrorRTrig(CLK := #System.Error);
       #PauseRTrig(CLK := #System.PauseOrders OR NOT #System.Auto_Man);
       IF #ErrorRTrig.Q OR #PauseRTrig.Q THEN
           #System.PauseOrders := FALSE;
           #System.Paused := #MaxRunningOrderNo > 0;
           IF #System.Paused THEN
               FOR #i := 1 TO UDINT_TO_DINT(#MaxRunningOrderNo) DO
                   IF #System.OrderTable[#i].Status = '' THEN
                       EXIT;
                   ELSIF #System.OrderTable[#i].Status = #QUEUED_STATUS THEN
                       #System.OrderTable[#i].Status := #PAUSED_STATUS;
                   ELSIF #System.OrderTable[#i].Status = #RUNNING_STATUS AND NOT #System.Auto_Man THEN
                       #System.OrderTable[#i].Status := #CANCELED_STATUS;
                   END_IF;
               END_FOR;
           END_IF;
       END_IF;
       IF #System.Paused AND #MaxRunningOrderNo = 0 THEN
           #System.Paused := FALSE;
       END_IF;
   END_REGION

   REGION Cancel Orders
       #CancelRTrig(CLK := #System.CancelOrders);
       #WeighingStation.Cancel := #ProfileStation.Cancel := #CancelRTrig.Q;
       IF #CancelRTrig.Q THEN
           #Canceling := TRUE;
           #System.CancelOrders := FALSE;
           #System.Paused := FALSE;
           FOR #i := 1 TO UDINT_TO_DINT(#MaxRunningOrderNo) DO
               IF #System.OrderTable[#i].Status = '' THEN
                   CONTINUE;
               ELSIF #System.OrderTable[#i].Status = #PAUSED_STATUS
                   OR #System.OrderTable[#i].Status = #QUEUED_STATUS
               THEN
                   #System.OrderTable[#i].Status := #CANCELED_STATUS;
                   #System.OrderTable[#i].CompleteTime := #CurrentTime;
               ELSIF #System.OrderTable[#i].Status = #ERROR_STATUS
               THEN
                   #System.OrderTable[#i].Status := #ERROR_CANCELED_STATUS;
                   #System.OrderTable[#i].CompleteTime := #CurrentTime;
               END_IF;
           END_FOR;
           #System.CurrentOrder := 0;
       END_IF;
       IF #Canceling AND NOT (#Cnv_Entry.Running OR #Cnv_PopUp_1.Running OR #WeighingStation.Running OR #ProfileStation.Running
           OR #Cnv_PopUp_2.Running OR #Cnv_PopUp_3.Running OR #Cnv_PopUp_4.Running OR #Cnv_Exit.Running) THEN
           #Canceling := FALSE;
           #Roller_To_Roller_CurrentOrder := #Chain_To_Chain_CurrentOrder:= #PickSt_To_Pop1_CurrentOrder := #Pop4_To_PickSt_CurrentOrder := 0;
            #WeighingStation_CurrentOrder:= #ProfileStation_CurrentOrder := 0;
       END_IF;
   END_REGION

   REGION Resume Orders
       #ResumeRTrig(CLK := #System.ResumeOrders);
       IF #ResumeRTrig.Q THEN
           #System.ResumeOrders := FALSE;
           #System.CurrentOrder := #MaxRunningOrderNo;
           IF NOT #System.Error THEN
               #System.Paused := FALSE;
               FOR #i := 1 TO UDINT_TO_DINT(#MaxRunningOrderNo) DO
                   IF #System.OrderTable[#i].Status = '' THEN
                       EXIT;
                   ELSIF #System.OrderTable[#i].Status = #PAUSED_STATUS
                       OR #System.OrderTable[#i].Status = #ERROR_STATUS
                   THEN
                       #System.OrderTable[#i].Status := #QUEUED_STATUS;
                   END_IF;
               END_FOR;
           END_IF;

       END_IF;
   END_REGION

   REGION Order Handler
       IF #System.Running AND NOT #System.Error
           AND (#System.OrderTable[#System.CurrentOrder].Status = #COMPLETED_STATUS
           OR #System.OrderTable[#System.CurrentOrder].Status = #ERROR_STATUS
           OR #System.OrderTable[#System.CurrentOrder].Status = #ERROR_CANCELED_STATUS
           OR #System.OrderTable[#System.CurrentOrder].Sequence = 0)
       THEN
           IF #System.CurrentOrder > 0 THEN
               #System.CurrentOrder -= 1;
           ELSE
               #System.CurrentOrder := 0;
           END_IF;
       END_IF;
   END_REGION

   REGION Watchdogs
       //Watchdog Timers
       #PickSt_To_Pop1WatchdogTimer(IN := #PickSt_To_Pop1WatchdogStart,
                                    PT := UDINT_TO_TIME(#Watchdog.Pick_TO_Pop1 * 60000),
                                    Q => #System.Watchdog_TimeOut.Pick_TO_Pop1);
       #Roller_To_Roller_WatchdogTimer(IN := #Roller_To_Roller_WatchdogStart,
                                       PT := UDINT_TO_TIME(#Watchdog.Roller_TO_Roller * 60000),
                                       Q => #System.Watchdog_TimeOut.Roller_TO_Roller);
       #Chain_To_Chain_WatchdogTimer(IN := #Chain_To_Chain_WatchdogStart,
                                     PT := UDINT_TO_TIME(#Watchdog.Chain_TO_Chain * 60000),
                                     Q => #System.Watchdog_TimeOut.Chain_TO_Chain);
       #Pop4_To_PickWatchdogTimer(IN := #Pop4_To_PickWatchdogStart,
                                  PT := UDINT_TO_TIME(#Watchdog.Pop4_TO_Pick * 60000),
                                  Q => #System.Watchdog_TimeOut.Pop4_TO_Pick);
       #WeighingStation_WatchdogTimer(IN := #WeighingStation_WatchdogStart,
                                      PT := UDINT_TO_TIME(#Watchdog.Weigh_Station * 60000),
                                      Q => #System.Watchdog_TimeOut.Weigh_Station);
       #ProfileStation_WatchdogTimer(IN := #ProfileStation_WatchdogStart,
                                     PT := UDINT_TO_TIME(#Watchdog.Profile_Station * 60000),
                                     Q => #System.Watchdog_TimeOut.Profile_Station);

       //Reset  Watchdog Timers
       IF #System.Error OR #CancelRTrig.Q OR #PauseRTrig.Q OR "Reset_All" THEN
           #PickSt_To_Pop1WatchdogStart := FALSE;
           #Roller_To_Roller_WatchdogStart := FALSE;
           #Chain_To_Chain_WatchdogStart := FALSE;
           #Pop4_To_PickWatchdogStart := FALSE;
           #WeighingStation_WatchdogStart := FALSE;
           #ProfileStation_WatchdogStart := FALSE;

       END_IF;
   END_REGION

   REGION Reset Next Order Number
       IF #System.NextOrder > 1
           AND #CurrentDTL.HOUR = 0
           AND #CurrentDTL.MINUTE = 0
           AND #CurrentDTL.SECOND = 0
       THEN
           #System.NextOrder := 1;
       END_IF;

   END_REGION

   REGION #System Mode and State
       #System.Selected := #System_Selected; // System selected
       #System.Ready := NOT #System.Error AND #System.Selected;
       #System.Auto_Man := #AutoMan_Switch;
       #System.Running := #Cnv_Entry.Running OR #Cnv_PopUp_1.Running OR #WeighingStation.Running
       OR #ProfileStation.Running OR #Cnv_PopUp_3.Running OR #Cnv_PopUp_4.Running;

       #System.Error := #Cnv_Entry.Error OR #Cnv_PopUp_1.Error OR #Cnv_PopUp_2.Error OR #Cnv_PopUp_3.Error OR #Cnv_PopUp_4.Error
       OR #Cnv_Exit.Error ; (*Implement Weigh station error and Profile Station error*)
       #System.IDLE := NOT #System.Running AND NOT #System.Paused AND NOT #System.Error;
       IF #System.Running THEN
           #System.State := 1;
       ELSIF #System.Paused AND NOT #System.Error THEN
           #System.State := 2;
       ELSIF #System.Error THEN
           #System.State := 3;
       ELSE
           #System.State := 0;
       END_IF;
   END_REGION
END_FUNCTION_BLOCK

FUNCTION_BLOCK "Order_Table_FB_VTD"   // FB31, SCL
{ S7_Optimized_Access := 'TRUE' }
VERSION : 0.1
// stored: AutoNumber false, IsIECCheckEnabled false, IsRetainMemResEnabled false, MemoryReserve 100, SetENOAutomatically false, UDAEnableTagReadback false
   VAR_INPUT
      System_Selected { ExternalWritable := 'False'} : Bool;
      AutoMan_Switch : Bool;   // Auto/Man Switch on CPU Panel - 1 = Auto, 0 = Manual
      CurrentTime { ExternalWritable := 'False'} : String;
      CurrentDTL : DTL;
      Watchdog : "Watchdog_Settings_UDT";
   END_VAR
   VAR_IN_OUT
      VTD : "VTD_Control";
      Extrator_Conveyor : "ECnv_Control";
      Cnv_Buffer_1 : "Buffer_Cnv_Control";
      Cnv_Buffer_2 : "Buffer_Cnv_Control";
      Cnv_Buffer_3 : "Buffer_Cnv_Control";
      System : "System_UDT";
      Control_OPC_Ua : "WMS_OPC_UA";
   END_VAR
   VAR
      VTD_CurrentOrder { ExternalWritable := 'False'} : UDInt := 0;
      Pallet_InOut_CurrentOrder : UDInt;
      Shuttle_InOut_CurrentOrder : UDInt;
      VTDDoneRTrig : R_TRIG;
      Pallet_InOut_RTrig { S7_SetPoint := 'True'} : R_TRIG;
      Shuttle_InOut_RTrig { S7_SetPoint := 'True'} : R_TRIG;
      PalletRefused_RTrig { ExternalWritable := 'False'} : R_TRIG;
      ErrorRTrig { ExternalWritable := 'False'} : R_TRIG;
      CancelRTrig { ExternalWritable := 'False'} : R_TRIG;
      PauseRTrig { ExternalWritable := 'False'} : R_TRIG;
      ResumeRTrig { ExternalWritable := 'False'} : R_TRIG;
      Clear_Store : R_TRIG;
      Clear_Retrieve : R_TRIG;
      Canceling : Bool;
      VTD_WatchdogTimer : TON_TIME;
      Pallet_InOut_WatchdogTimer { S7_SetPoint := 'True'} : TON_TIME;
      Shuttle_InOut_WatchdogTimer { S7_SetPoint := 'True'} : TON_TIME;
      VTD_WatchdogStart : Bool;
      Pallet_InOut_WatchdogStart : Bool;
      Shuttle_InOut_WatchdogStart : Bool;
   END_VAR
   VAR_TEMP
      i : DInt;
      n : DInt;
      EmptyOrder : "OrderTable_UDT";
      MaxRunningOrderNo : UInt;
   END_VAR
   VAR CONSTANT
      VTD_DEVICE : String := 'VTD';
      PALLET_INOUT_DEVICE : String := 'Pallet In Out';
      SHUTTLE_INOUT_DEVICE : String := 'Shuttle In Out';
      RUNNING_STATUS : String := 'Running';
      COMPLETED_STATUS : String := 'Completed';
      QUEUED_STATUS : String := 'Queued';
      PALLET_REFUSED_STATUS : String := 'Pallet Refused';
      ERROR_STATUS : String := 'Error';
      CANCELED_STATUS : String := 'Canceled';
      PAUSED_STATUS : String := 'Paused';
      ORDER_REFUSED : String := 'Refused';
      ERROR_CANCELED_STATUS : String := 'Error\Cancel';
   END_VAR
BEGIN

   // Converts the task type for strings 
   IF #System.OrderTable[1].OPC_Control.Task_Type = 1 THEN
       #System.OrderTable[1].Device := 'VTD';
   ELSIF #System.OrderTable[1].OPC_Control.Task_Type = 4 OR #System.OrderTable[1].OPC_Control.Task_Type = 5  THEN
       #System.OrderTable[1].Device := 'Pallet In Out';
   ELSIF #System.OrderTable[1].OPC_Control.Task_Type = 2 OR #System.OrderTable[1].OPC_Control.Task_Type = 3 THEN
       #System.OrderTable[1].Device := 'Shuttle In Out';
   ELSE
       #System.OrderTable[1].Device := '';
   END_IF;


   REGION #New Order was Sent
       IF #System.OrderSent THEN
           //Count orders in Step Table
           FOR #i := 0 TO 20 DO
               IF #System.StepTable[#i].OrderNo <> 0
                   AND #System.StepTable[#i].StepNo <> 0
                   AND #System.StepTable[#i].PlaceTime <> ''
                   //AND #System.StepTable[#i].Device <> ''
                   AND #System.StepTable[#i].Status = #QUEUED_STATUS
               THEN
                   #n += 1;
               ELSE
                   EXIT;
               END_IF;
           END_FOR;
           IF #n > 0 THEN
               //shift order table down by Order number rows
               FOR #i := 99 TO (#n + 1) BY -1 DO
                   #System.OrderTable[#i] := #System.OrderTable[#i - #n];
               END_FOR;
               //copy data from step table to order table
               FOR #i := 0 (*1*) TO #n DO
                   #System.OrderTable[#n - #i (*+ 1*)] := #System.StepTable[#i];
               END_FOR;
               //clean step table
               FOR #i := 0 (*1*) TO 20 DO
                   #System.StepTable[#i] := #EmptyOrder;
               END_FOR;
               #System.CurrentOrder += #n;

               //VTD move to floor
               IF #VTD_CurrentOrder <> 0 THEN
                   #VTD_CurrentOrder += #n;
               END_IF;

               //Shuttle transfer in/out of the VTD
               IF #Pallet_InOut_CurrentOrder <> 0 THEN
                   #Pallet_InOut_CurrentOrder += #n;
               END_IF;

               //Transfer Pallet in/out of the VTD
               IF #Shuttle_InOut_CurrentOrder <> 0 THEN
                   #Shuttle_InOut_CurrentOrder += #n;
               END_IF;

                       END_IF;
           #System.OrderSent := FALSE;
       END_IF;
   END_REGION

   REGION Auto/Man Mode
       //Enable Devices in Auto/Man Mode
       IF #System.Auto_Man THEN
          // #VTD.Mode := #Extrator_Conveyor.Mode := #Cnv_Buffer_1.Mode := #Cnv_Buffer_2.Mode := #Cnv_Buffer_3.Mode := 3;// Auto Mode
           #VTD.Instruction.Enable := #Extrator_Conveyor.Enabled := #Cnv_Buffer_1.Instruction.Enable :=
           #Cnv_Buffer_2.Instruction.Enable := #Cnv_Buffer_3.Instruction.Enable := TRUE; // := Not System.Error
       ELSE //Disable Devices in Auto/Man Mode

           //#VTD.Mode := #Extrator_Conveyor.Mode := #Cnv_Buffer_1.Mode := #Cnv_Buffer_2.Mode := #Cnv_Buffer_3.Mode := 0;
           #VTD.Instruction.Enable := #Extrator_Conveyor.Enabled := #Cnv_Buffer_1.Instruction.Enable :=
           #Cnv_Buffer_2.Instruction.Enable := #Cnv_Buffer_3.Instruction.Enable := FALSE;
       END_IF;
   END_REGION

   REGION VTD
       //VTD 
       IF #System.OrderTable[1].StepNo <> 0
           AND #System.OrderTable[1].Device = #VTD_DEVICE
           AND #System.OrderTable[1].Status = #QUEUED_STATUS
           AND NOT ("OPC_UA_Control_FB_DB".State_VTD > 20 AND "OPC_UA_Control_FB_DB".State_VTD < 400)
           AND NOT #System.Error
           AND NOT #Canceling
       THEN
           #VTD_CurrentOrder := 1;
       END_IF;
       IF #System.OrderTable[#VTD_CurrentOrder].StepNo <> 0
           AND #System.OrderTable[#VTD_CurrentOrder].Device = #VTD_DEVICE
           AND #System.OrderTable[#VTD_CurrentOrder].Status = #QUEUED_STATUS
           AND NOT ("OPC_UA_Control_FB_DB".State_VTD > 20 AND "OPC_UA_Control_FB_DB".State_VTD < 400)
           AND NOT #System.Error
           AND NOT #Canceling
       THEN

           //OPC Commands to Move VTD between floors
           // WCS => Order Table => OPC Ua Control Table

           "Control_DB"."VTD_Order Table".Task_Data_Available:= TRUE;//#System.OrderTable[#VTD_CurrentOrder].OPC_Control.Task_Data_Available; // Send the Task Data Available from WCS 
           "Control_DB"."VTD_Order Table".Task_Type:= #System.OrderTable[#VTD_CurrentOrder].OPC_Control.Task_Type; // Send the Task Type - VTD = Task Type = 1
           "Control_DB"."VTD_Order Table".Pallet_Type:= #System.OrderTable[#VTD_CurrentOrder].OPC_Control.Pallet_Type; // Send the Pallet Type -C=Chep/E=Euro
           "Control_DB"."VTD_Order Table".Task_ID:=#System.OrderTable[#VTD_CurrentOrder].OPC_Control.Task_ID; // Send the Task ID number;
           "Control_DB"."VTD_Order Table".Task_Metadata:=#System.OrderTable[#VTD_CurrentOrder].OPC_Control.Task_Metadata; // Send the Task Metadata Unique identifier
           "Control_DB"."VTD_Order Table".Destination_Location:= #System.OrderTable[#VTD_CurrentOrder].OPC_Control.Destination_Location; // Send the VTD Destination Location
           "Control_DB"."VTD_Order Table".Source_Location := 0; // Send the VTD Destination Location
           #VTD_WatchdogStart := TRUE;
       END_IF;

       //RUNNING
       IF ("OPC_UA_Control_FB_DB".State_VTD > 20 AND "OPC_UA_Control_FB_DB".State_VTD < 400) AND #System.Auto_Man THEN
           //#VTD.Instruction.Execulte := FALSE;
           #System.OrderTable[#VTD_CurrentOrder].Status := #RUNNING_STATUS;
            "Control_DB"."VTD_Order Table".Task_Data_Available := FALSE; // Send the Task Data Available from WCS 
           // "Control_DB"."VTD_Order Table".Task_Type := 0; // Send the Task Type - VTD = Task Type = 1
           // "Control_DB"."VTD_Order Table".Pallet_Type := ' '; // Send the Pallet Type -C=Chep/E=Euro
           // "Control_DB"."VTD_Order Table".Task_ID := 0; // Send the Task ID number;
           // "Control_DB"."VTD_Order Table".Task_Metadata := ''; // Send the Task Metadata Unique identifier
           // "Control_DB"."VTD_Order Table".Destination_Location := 0; // Send the VTD Destination Location
           // "Control_DB"."VTD_Order Table".Source_Location := 0; // Send the VTD Destination Location

       END_IF;

       //Cancel order
       IF #Canceling AND NOT #VTD.Running AND #VTD_CurrentOrder <> 0 THEN
           #System.OrderTable[#VTD_CurrentOrder].Status := #CANCELED_STATUS;
           #System.OrderTable[#VTD_CurrentOrder].CompleteTime := #CurrentTime;
           #VTD_CurrentOrder := 0;
          // #VTD.Instruction.Execulte := FALSE;
           "Control_DB"."VTD_Order Table".Task_Data_Available := FALSE; // Send the Task Data Available from WCS 
           "Control_DB"."VTD_Order Table".Task_Type := 0; // Send the Task Type - VTD = Task Type = 1
           "Control_DB"."VTD_Order Table".Pallet_Type := ' '; // Send the Pallet Type -C=Chep/E=Euro
           "Control_DB"."VTD_Order Table".Task_ID := 0; // Send the Task ID number;
           "Control_DB"."VTD_Order Table".Task_Metadata := ''; // Send the Task Metadata Unique identifier
           "Control_DB"."VTD_Order Table".Destination_Location := 0; // Send the VTD Destination Location
           "Control_DB"."VTD_Order Table".Source_Location := 0; // Send the VTD Destination 
       END_IF;

       //Error
       IF #VTD.Error THEN
           //#VTD.Instruction.Execulte := FALSE;
           "Control_DB"."VTD_Order Table".Task_Data_Available := FALSE; // Send the Task Data Available from WCS 
           "Control_DB"."VTD_Order Table".Task_Type := 0; // Send the Task Type - VTD = Task Type = 1
           "Control_DB"."VTD_Order Table".Pallet_Type := ' '; // Send the Pallet Type -C=Chep/E=Euro
           "Control_DB"."VTD_Order Table".Task_ID := 0; // Send the Task ID number;
           "Control_DB"."VTD_Order Table".Task_Metadata := ''; // Send the Task Metadata Unique identifier
           "Control_DB"."VTD_Order Table".Destination_Location := 0; // Send the VTD Destination Location
           "Control_DB"."VTD_Order Table".Source_Location := 0; // Send the VTD Destination 
           #System.OrderTable[#VTD_CurrentOrder].ErrorID := #VTD.VTD_Errors.Error_Word_1;
       END_IF;

       //MOVEMENT FINALIZED
       #VTDDoneRTrig(CLK := "Control_DB"."VTD_Order Table".Movement_Request_Complete );
       IF #VTDDoneRTrig.Q THEN
           // "Control_DB"."VTD_Order Table".Task_Data_Available := FALSE; // Send the Task Data Available from WCS 
           // "Control_DB"."VTD_Order Table".Task_Type := 0; // Send the Task Type - VTD = Task Type = 1
           // "Control_DB"."VTD_Order Table".Pallet_Type := ' '; // Send the Pallet Type -C=Chep/E=Euro
           // "Control_DB"."VTD_Order Table".Task_ID := 0; // Send the Task ID number;
           // "Control_DB"."VTD_Order Table".Task_Metadata := ''; // Send the Task Metadata Unique identifier
           // "Control_DB"."VTD_Order Table".Destination_Location := 0; // Send the VTD Destination Location
           // "Control_DB"."VTD_Order Table".Source_Location := 0; // Send the VTD Destination 
           #VTD_WatchdogStart := FALSE;
           #System.OrderTable[#VTD_CurrentOrder].Status := #COMPLETED_STATUS;
           #System.OrderTable[#VTD_CurrentOrder].CompleteTime := #CurrentTime;
           #VTD_CurrentOrder := 0;
       END_IF;
   END_REGION
   ///////////////////////////////////////////////////////////////////////////////////////////////////////////////////////////////////////
   ///////////////////////////////////////////////////////////////////////////////////////////////////////////////////////////////////////
   REGION Pallet_InOut - Conveyors
       //VTD 
       IF #System.OrderTable[1].StepNo <> 0
           AND #System.OrderTable[1].Device = #PALLET_INOUT_DEVICE
           AND #System.OrderTable[1].Status = #QUEUED_STATUS
           AND NOT ("OPC_UA_Control_FB_DB".State_VTD > 20 AND "OPC_UA_Control_FB_DB".State_VTD < 400)
           AND NOT #System.Error
           AND NOT #Canceling
       THEN
           #Pallet_InOut_CurrentOrder := 1;
       END_IF;
       IF #System.OrderTable[#Pallet_InOut_CurrentOrder].StepNo <> 0
           AND #System.OrderTable[#Pallet_InOut_CurrentOrder].Device = #PALLET_INOUT_DEVICE
           AND #System.OrderTable[#Pallet_InOut_CurrentOrder].Status = #QUEUED_STATUS
           AND NOT ("OPC_UA_Control_FB_DB".State_VTD > 20 AND "OPC_UA_Control_FB_DB".State_VTD < 400)
           AND NOT #System.Error
           AND NOT #Canceling
       THEN
           //OPC Commands to Move Pallets IN/OUT (Buffer conveyors/Extractor conveyors)
           // WCS => Order Table => OPC Ua Control Table
           "Control_DB"."VTD_Order Table".Task_Data_Available := TRUE; //#System.OrderTable[#Pallet_InOut_CurrentOrder].OPC_Control.Task_Data_Available; // Send the Task Data Available from WCS 
           "Control_DB"."VTD_Order Table".Task_Type := #System.OrderTable[#Pallet_InOut_CurrentOrder].OPC_Control.Task_Type; // Send the Task Type - Pallet Transfer IN/OUT = Task Type = 4/
           "Control_DB"."VTD_Order Table".Task_ID := #System.OrderTable[#Pallet_InOut_CurrentOrder].OPC_Control.Task_ID; // Send the Task ID number;
           "Control_DB"."VTD_Order Table".Task_Metadata := #System.OrderTable[#Pallet_InOut_CurrentOrder].OPC_Control.Task_Metadata; // Send the Task Metadata Unique identifier
           "Control_DB"."VTD_Order Table".Source_Location := #System.OrderTable[#Pallet_InOut_CurrentOrder].OPC_Control.Source_Location; // Send the Source Location from the Conveyor
           "Control_DB"."VTD_Order Table".Destination_Location := #System.OrderTable[#Pallet_InOut_CurrentOrder].OPC_Control.Destination_Location; // Send the Destination Location to the Conveyor;
           #Pallet_InOut_WatchdogStart := TRUE;
       END_IF;

       //RUNNING
       IF (#Cnv_Buffer_1.Running OR #Cnv_Buffer_2.Running OR #Cnv_Buffer_3.Running OR #Extrator_Conveyor.Running) AND #System.Auto_Man THEN
          // #VTD.Instruction.Execulte := FALSE;
           #System.OrderTable[#Pallet_InOut_CurrentOrder].Status := #RUNNING_STATUS;
           // "Control_DB"."VTD_Order Table".Task_Data_Available := FALSE; //#System.OrderTable[#Pallet_InOut_CurrentOrder].OPC_Control.Task_Data_Available; // Send the Task Data Available from WCS 
           // "Control_DB"."VTD_Order Table".Task_Type := #System.OrderTable[#Pallet_InOut_CurrentOrder].OPC_Control.Task_Type; // Send the Task Type - Pallet Transfer IN/OUT = Task Type = 4/
           // "Control_DB"."VTD_Order Table".Task_ID := #System.OrderTable[#Pallet_InOut_CurrentOrder].OPC_Control.Task_ID; // Send the Task ID number;
           // "Control_DB"."VTD_Order Table".Task_Metadata := #System.OrderTable[#Pallet_InOut_CurrentOrder].OPC_Control.Task_Metadata; // Send the Task Metadata Unique identifier
           // "Control_DB"."VTD_Order Table".Source_Location := #System.OrderTable[#Pallet_InOut_CurrentOrder].OPC_Control.Source_Location; // Send the Source Location from the Conveyor
           // "Control_DB"."VTD_Order Table".Destination_Location := #System.OrderTable[#Pallet_InOut_CurrentOrder].OPC_Control.Destination_Location; // Send the Destination Location to the Conveyor;

       END_IF;

       //Cancel order
       IF #Canceling AND NOT (#Cnv_Buffer_1.Running OR #Cnv_Buffer_2.Running OR #Cnv_Buffer_3.Running OR #Extrator_Conveyor.Running) AND #Pallet_InOut_CurrentOrder <> 0 THEN
           #System.OrderTable[#Pallet_InOut_CurrentOrder].Status := #CANCELED_STATUS;
           #System.OrderTable[#Pallet_InOut_CurrentOrder].CompleteTime := #CurrentTime;
           #Pallet_InOut_CurrentOrder := 0;
           //#VTD.Instruction.Execulte := FALSE;
           //
           "Control_DB"."VTD_Order Table".Task_Data_Available := FALSE; //#System.OrderTable[#Pallet_InOut_CurrentOrder].OPC_Control.Task_Data_Available; // Send the Task Data Available from WCS 
           "Control_DB"."VTD_Order Table".Task_Type := #System.OrderTable[#Pallet_InOut_CurrentOrder].OPC_Control.Task_Type; // Send the Task Type - Pallet Transfer IN/OUT = Task Type = 4/
           "Control_DB"."VTD_Order Table".Task_ID := #System.OrderTable[#Pallet_InOut_CurrentOrder].OPC_Control.Task_ID; // Send the Task ID number;
           "Control_DB"."VTD_Order Table".Task_Metadata := #System.OrderTable[#Pallet_InOut_CurrentOrder].OPC_Control.Task_Metadata; // Send the Task Metadata Unique identifier
           "Control_DB"."VTD_Order Table".Source_Location := #System.OrderTable[#Pallet_InOut_CurrentOrder].OPC_Control.Source_Location; // Send the Source Location from the Conveyor
           "Control_DB"."VTD_Order Table".Destination_Location := #System.OrderTable[#Pallet_InOut_CurrentOrder].OPC_Control.Destination_Location; // Send the Destination Location to the Conveyor;

       END_IF;

       //Error

       IF (#Cnv_Buffer_1.Error OR #Cnv_Buffer_2.Error OR #Cnv_Buffer_3.Error OR #Extrator_Conveyor.Error) THEN
           // #VTD.Instruction.Execulte := FALSE;
           "Control_DB"."VTD_Order Table".Task_Data_Available := FALSE; //#System.OrderTable[#Pallet_InOut_CurrentOrder].OPC_Control.Task_Data_Available; // Send the Task Data Available from WCS 
           "Control_DB"."VTD_Order Table".Task_Type := #System.OrderTable[#Pallet_InOut_CurrentOrder].OPC_Control.Task_Type; // Send the Task Type - Pallet Transfer IN/OUT = Task Type = 4/
           "Control_DB"."VTD_Order Table".Task_ID := #System.OrderTable[#Pallet_InOut_CurrentOrder].OPC_Control.Task_ID; // Send the Task ID number;
           "Control_DB"."VTD_Order Table".Task_Metadata := #System.OrderTable[#Pallet_InOut_CurrentOrder].OPC_Control.Task_Metadata; // Send the Task Metadata Unique identifier
           "Control_DB"."VTD_Order Table".Source_Location := #System.OrderTable[#Pallet_InOut_CurrentOrder].OPC_Control.Source_Location; // Send the Source Location from the Conveyor
           "Control_DB"."VTD_Order Table".Destination_Location := #System.OrderTable[#Pallet_InOut_CurrentOrder].OPC_Control.Destination_Location; // Send the Destination Location to the Conveyor;

           #System.OrderTable[#Pallet_InOut_CurrentOrder].ErrorID := (#Cnv_Buffer_1.Cnv_Errors.Error_Word_1
                                                                   OR #Cnv_Buffer_2.Cnv_Errors.Error_Word_1
                                                                   OR #Cnv_Buffer_3.Cnv_Errors.Error_Word_1
                                                                   OR #Extrator_Conveyor.Cnv_Errors.Error_Word_1);
       END_IF;

       //MOVEMENT FINALIZED
       #Pallet_InOut_RTrig(CLK := "Control_DB"."VTD_Order Table".Movement_Request_Complete);
       IF #Pallet_InOut_RTrig.Q THEN

           "Control_DB"."VTD_Order Table".Task_Data_Available := FALSE; //#System.OrderTable[#Pallet_InOut_CurrentOrder].OPC_Control.Task_Data_Available; // Send the Task Data Available from WCS 
           "Control_DB"."VTD_Order Table".Task_Type := #System.OrderTable[#Pallet_InOut_CurrentOrder].OPC_Control.Task_Type; // Send the Task Type - Pallet Transfer IN/OUT = Task Type = 4/
           "Control_DB"."VTD_Order Table".Task_ID := #System.OrderTable[#Pallet_InOut_CurrentOrder].OPC_Control.Task_ID; // Send the Task ID number;
           "Control_DB"."VTD_Order Table".Task_Metadata := #System.OrderTable[#Pallet_InOut_CurrentOrder].OPC_Control.Task_Metadata; // Send the Task Metadata Unique identifier
           "Control_DB"."VTD_Order Table".Source_Location := #System.OrderTable[#Pallet_InOut_CurrentOrder].OPC_Control.Source_Location; // Send the Source Location from the Conveyor
           "Control_DB"."VTD_Order Table".Destination_Location := #System.OrderTable[#Pallet_InOut_CurrentOrder].OPC_Control.Destination_Location; // Send the Destination Location to the Conveyor;

           #System.OrderTable[#Pallet_InOut_CurrentOrder].Status := #COMPLETED_STATUS;
           #System.OrderTable[#Pallet_InOut_CurrentOrder].CompleteTime := #CurrentTime;
           #Pallet_InOut_CurrentOrder := 0;
       END_IF;
   END_REGION
   ///////////////////////////////////////////////////////////////////////////////////////////////////////////////////////////////////////
   ///////////////////////////////////////////////////////////////////////////////////////////////////////////////////////////////////////
   REGION Shuttle_InOut
       //Shuttle Interlock on VTD 
       IF #System.OrderTable[1].StepNo <> 0
           AND #System.OrderTable[1].Device = #SHUTTLE_INOUT_DEVICE
           AND #System.OrderTable[1].Status = #QUEUED_STATUS
           AND NOT ("OPC_UA_Control_FB_DB".State_VTD > 20 AND "OPC_UA_Control_FB_DB".State_VTD < 400)
           AND NOT #System.Error
           AND NOT #Canceling
       THEN
           #Shuttle_InOut_CurrentOrder := 1;
       END_IF;
       IF #System.OrderTable[#Shuttle_InOut_CurrentOrder].StepNo <> 0
           AND #System.OrderTable[#Shuttle_InOut_CurrentOrder].Device = #SHUTTLE_INOUT_DEVICE
           AND #System.OrderTable[#Shuttle_InOut_CurrentOrder].Status = #QUEUED_STATUS
           AND NOT ("OPC_UA_Control_FB_DB".State_VTD > 20 AND "OPC_UA_Control_FB_DB".State_VTD < 400)
           AND NOT #System.Error
           AND NOT #Canceling
       THEN
           //OPC Commands to Move Shuttle IN/OUT (Shuttles IN/OUT)
           // WCS => Order Table => OPC Ua Control Table

           "Control_DB"."VTD_Order Table".Task_Data_Available := TRUE;//#System.OrderTable[#Shuttle_InOut_CurrentOrder].OPC_Control.Task_Data_Available; // Send the Task Data Available from WCS 
           "Control_DB"."VTD_Order Table".Task_ID := #System.OrderTable[#Shuttle_InOut_CurrentOrder].OPC_Control.Task_ID; // Send the Task ID number;
           "Control_DB"."VTD_Order Table".Task_Metadata := #System.OrderTable[#Shuttle_InOut_CurrentOrder].OPC_Control.Task_Metadata; // Send the Task Metadata Unique identifier
           "Control_DB"."VTD_Order Table".Pallet_Type := #System.OrderTable[#Shuttle_InOut_CurrentOrder].OPC_Control.Pallet_Type; // Send Pallet Type
           "Control_DB"."VTD_Order Table".Task_Type := #System.OrderTable[#Shuttle_InOut_CurrentOrder].OPC_Control.Task_Type; // Send the Task Type - Pallet Transfer IN/OUT = Task Type = 4/
           "Control_DB"."VTD_Order Table".Shuttle_ID := #System.OrderTable[#Shuttle_InOut_CurrentOrder].OPC_Control.Shuttle_ID;// Send the Shuttle ID
           "Control_DB"."VTD_Order Table".Shuttle_Loaded := #System.OrderTable[#Shuttle_InOut_CurrentOrder].OPC_Control.Shuttle_Loaded; // Send the Shuttle status (Loaded/Unloaded)
           "Control_DB"."VTD_Order Table".Source_Location := #System.OrderTable[#Shuttle_InOut_CurrentOrder].OPC_Control.Source_Location; // Send the Source Location from the Conveyor
           "Control_DB"."VTD_Order Table".Destination_Location := #System.OrderTable[#Shuttle_InOut_CurrentOrder].OPC_Control.Destination_Location; // Send the Destination Location to the Conveyor;
           #Shuttle_InOut_WatchdogStart := TRUE;
       END_IF;

       //RUNNING
       IF (#VTD.Running) AND #System.Auto_Man THEN
           //#VTD.Instruction.Execulte := FALSE;
           #System.OrderTable[#Shuttle_InOut_CurrentOrder].Status := #RUNNING_STATUS;
           // "Control_DB"."VTD_Order Table".Task_Data_Available := FALSE;//#System.OrderTable[#Shuttle_InOut_CurrentOrder].OPC_Control.Task_Data_Available; // Send the Task Data Available from WCS 
           // "Control_DB"."VTD_Order Table".Task_ID := #System.OrderTable[#Shuttle_InOut_CurrentOrder].OPC_Control.Task_ID; // Send the Task ID number;
           // "Control_DB"."VTD_Order Table".Task_Metadata := #System.OrderTable[#Shuttle_InOut_CurrentOrder].OPC_Control.Task_Metadata; // Send the Task Metadata Unique identifier
           // "Control_DB"."VTD_Order Table".Pallet_Type := #System.OrderTable[#Shuttle_InOut_CurrentOrder].OPC_Control.Pallet_Type; // Send Pallet Type
           // "Control_DB"."VTD_Order Table".Task_Type := #System.OrderTable[#Shuttle_InOut_CurrentOrder].OPC_Control.Task_Type; // Send the Task Type - Pallet Transfer IN/OUT = Task Type = 4/
           // "Control_DB"."VTD_Order Table".Shuttle_ID := #System.OrderTable[#Shuttle_InOut_CurrentOrder].OPC_Control.Shuttle_ID;// Send the Shuttle ID
           // "Control_DB"."VTD_Order Table".Shuttle_Loaded := #System.OrderTable[#Shuttle_InOut_CurrentOrder].OPC_Control.Shuttle_Loaded; // Send the Shuttle status (Loaded/Unloaded)
           // "Control_DB"."VTD_Order Table".Source_Location := #System.OrderTable[#Shuttle_InOut_CurrentOrder].OPC_Control.Source_Location; // Send the Source Location from the Conveyor
           // "Control_DB"."VTD_Order Table".Destination_Location := #System.OrderTable[#Shuttle_InOut_CurrentOrder].OPC_Control.Destination_Location; // Send the Destination Location to the Conveyor;

       END_IF;

       //Cancel order
       IF #Canceling AND NOT (#VTD.Running) AND #Shuttle_InOut_CurrentOrder <> 0 THEN
           #System.OrderTable[#Shuttle_InOut_CurrentOrder].Status := #CANCELED_STATUS;
           #System.OrderTable[#Shuttle_InOut_CurrentOrder].CompleteTime := #CurrentTime;
           #Shuttle_InOut_CurrentOrder := 0;
           //#VTD.Instruction.Execulte := FALSE;
           "Control_DB"."VTD_Order Table".Task_Data_Available := FALSE;//#System.OrderTable[#Shuttle_InOut_CurrentOrder].OPC_Control.Task_Data_Available; // Send the Task Data Available from WCS 
           "Control_DB"."VTD_Order Table".Task_ID := #System.OrderTable[#Shuttle_InOut_CurrentOrder].OPC_Control.Task_ID; // Send the Task ID number;
           "Control_DB"."VTD_Order Table".Task_Metadata := #System.OrderTable[#Shuttle_InOut_CurrentOrder].OPC_Control.Task_Metadata; // Send the Task Metadata Unique identifier
           "Control_DB"."VTD_Order Table".Pallet_Type := #System.OrderTable[#Shuttle_InOut_CurrentOrder].OPC_Control.Pallet_Type; // Send Pallet Type
           "Control_DB"."VTD_Order Table".Task_Type := #System.OrderTable[#Shuttle_InOut_CurrentOrder].OPC_Control.Task_Type; // Send the Task Type - Pallet Transfer IN/OUT = Task Type = 4/
           "Control_DB"."VTD_Order Table".Shuttle_ID := #System.OrderTable[#Shuttle_InOut_CurrentOrder].OPC_Control.Shuttle_ID;// Send the Shuttle ID
           "Control_DB"."VTD_Order Table".Shuttle_Loaded := #System.OrderTable[#Shuttle_InOut_CurrentOrder].OPC_Control.Shuttle_Loaded; // Send the Shuttle status (Loaded/Unloaded)
           "Control_DB"."VTD_Order Table".Source_Location := #System.OrderTable[#Shuttle_InOut_CurrentOrder].OPC_Control.Source_Location; // Send the Source Location from the Conveyor
           "Control_DB"."VTD_Order Table".Destination_Location := #System.OrderTable[#Shuttle_InOut_CurrentOrder].OPC_Control.Destination_Location; // Send the Destination Location to the Conveyor;

       END_IF;

       //Error

       IF (#VTD.Error) THEN
           // #VTD.Instruction.Execulte := FALSE;
           "Control_DB"."VTD_Order Table".Task_Data_Available := FALSE;//#System.OrderTable[#Shuttle_InOut_CurrentOrder].OPC_Control.Task_Data_Available; // Send the Task Data Available from WCS 
           "Control_DB"."VTD_Order Table".Task_ID := #System.OrderTable[#Shuttle_InOut_CurrentOrder].OPC_Control.Task_ID; // Send the Task ID number;
           "Control_DB"."VTD_Order Table".Task_Metadata := #System.OrderTable[#Shuttle_InOut_CurrentOrder].OPC_Control.Task_Metadata; // Send the Task Metadata Unique identifier
           "Control_DB"."VTD_Order Table".Pallet_Type := #System.OrderTable[#Shuttle_InOut_CurrentOrder].OPC_Control.Pallet_Type; // Send Pallet Type
           "Control_DB"."VTD_Order Table".Task_Type := #System.OrderTable[#Shuttle_InOut_CurrentOrder].OPC_Control.Task_Type; // Send the Task Type - Pallet Transfer IN/OUT = Task Type = 4/
           "Control_DB"."VTD_Order Table".Shuttle_ID := #System.OrderTable[#Shuttle_InOut_CurrentOrder].OPC_Control.Shuttle_ID;// Send the Shuttle ID
           "Control_DB"."VTD_Order Table".Shuttle_Loaded := #System.OrderTable[#Shuttle_InOut_CurrentOrder].OPC_Control.Shuttle_Loaded; // Send the Shuttle status (Loaded/Unloaded)
           "Control_DB"."VTD_Order Table".Source_Location := #System.OrderTable[#Shuttle_InOut_CurrentOrder].OPC_Control.Source_Location; // Send the Source Location from the Conveyor
           "Control_DB"."VTD_Order Table".Destination_Location := #System.OrderTable[#Shuttle_InOut_CurrentOrder].OPC_Control.Destination_Location; // Send the Destination Location to the Conveyor;

           #System.OrderTable[#Shuttle_InOut_CurrentOrder].ErrorID := (#VTD.VTD_Errors.Error_Word_3);
       END_IF;

       //MOVEMENT FINALIZED
       #Shuttle_InOut_RTrig(CLK := #VTD.Shuttle_Interlock.Interlock_Complete);
       IF #Shuttle_InOut_RTrig.Q THEN
           "Control_DB"."VTD_Order Table".Task_Data_Available := FALSE;//#System.OrderTable[#Shuttle_InOut_CurrentOrder].OPC_Control.Task_Data_Available; // Send the Task Data Available from WCS 
           "Control_DB"."VTD_Order Table".Task_ID := #System.OrderTable[#Shuttle_InOut_CurrentOrder].OPC_Control.Task_ID; // Send the Task ID number;
           "Control_DB"."VTD_Order Table".Task_Metadata := #System.OrderTable[#Shuttle_InOut_CurrentOrder].OPC_Control.Task_Metadata; // Send the Task Metadata Unique identifier
           "Control_DB"."VTD_Order Table".Pallet_Type := #System.OrderTable[#Shuttle_InOut_CurrentOrder].OPC_Control.Pallet_Type; // Send Pallet Type
           "Control_DB"."VTD_Order Table".Task_Type := #System.OrderTable[#Shuttle_InOut_CurrentOrder].OPC_Control.Task_Type; // Send the Task Type - Pallet Transfer IN/OUT = Task Type = 4/
           "Control_DB"."VTD_Order Table".Shuttle_ID := #System.OrderTable[#Shuttle_InOut_CurrentOrder].OPC_Control.Shuttle_ID;// Send the Shuttle ID
           "Control_DB"."VTD_Order Table".Shuttle_Loaded := #System.OrderTable[#Shuttle_InOut_CurrentOrder].OPC_Control.Shuttle_Loaded; // Send the Shuttle status (Loaded/Unloaded)
           "Control_DB"."VTD_Order Table".Source_Location := #System.OrderTable[#Shuttle_InOut_CurrentOrder].OPC_Control.Source_Location; // Send the Source Location from the Conveyor
           "Control_DB"."VTD_Order Table".Destination_Location := #System.OrderTable[#Shuttle_InOut_CurrentOrder].OPC_Control.Destination_Location; // Send the Destination Location to the Conveyor;

           #Shuttle_InOut_WatchdogStart := FALSE;
           #System.OrderTable[#Shuttle_InOut_CurrentOrder].Status := #COMPLETED_STATUS;
           #System.OrderTable[#Shuttle_InOut_CurrentOrder].CompleteTime := #CurrentTime;
           #Shuttle_InOut_CurrentOrder := 0;
       END_IF;
   END_REGION


   REGION Max Running Order Number
       #MaxRunningOrderNo := MAX(IN1 := #VTD_CurrentOrder, IN2 := #Pallet_InOut_CurrentOrder,
                                 IN3 := #Shuttle_InOut_CurrentOrder, IN4 := #System.CurrentOrder);

   END_REGION

   REGION Pause Orders
       #ErrorRTrig(CLK := #System.Error);
       #PauseRTrig(CLK := #System.PauseOrders OR NOT #System.Auto_Man);
       IF #ErrorRTrig.Q OR #PauseRTrig.Q THEN
           #System.PauseOrders := FALSE;
           #System.Paused := #MaxRunningOrderNo > 0;
           IF #System.Paused THEN
               FOR #i := 1 TO UDINT_TO_DINT(#MaxRunningOrderNo) DO
                   IF #System.OrderTable[#i].Status = '' THEN
                       EXIT;
                   ELSIF #System.OrderTable[#i].Status = #QUEUED_STATUS THEN
                       #System.OrderTable[#i].Status := #PAUSED_STATUS;
                   ELSIF #System.OrderTable[#i].Status = #RUNNING_STATUS AND NOT #System.Auto_Man THEN
                       #System.OrderTable[#i].Status := #CANCELED_STATUS;
                   END_IF;
               END_FOR;
           END_IF;
       END_IF;
       IF #System.Paused AND #MaxRunningOrderNo = 0 THEN
           #System.Paused := FALSE;
       END_IF;
   END_REGION

   REGION Cancel Orders
       #CancelRTrig(CLK := #System.CancelOrders);
       (*#WeighingStation.Cancel := #ProfileStation.Cancel:= #CancelRTrig.Q*);
       IF #CancelRTrig.Q THEN
           #Canceling := TRUE;
           #System.CancelOrders := FALSE;
           #System.Paused := FALSE;
           FOR #i := 1 TO UDINT_TO_DINT(#MaxRunningOrderNo) DO
               IF #System.OrderTable[#i].Status = '' THEN
                   CONTINUE;
               ELSIF #System.OrderTable[#i].Status = #PAUSED_STATUS
                   OR #System.OrderTable[#i].Status = #QUEUED_STATUS
               THEN
                   #System.OrderTable[#i].Status := #CANCELED_STATUS;
                   #System.OrderTable[#i].CompleteTime := #CurrentTime;
               ELSIF #System.OrderTable[#i].Status = #ERROR_STATUS
               THEN
                   #System.OrderTable[#i].Status := #ERROR_CANCELED_STATUS;
                   #System.OrderTable[#i].CompleteTime := #CurrentTime;
               END_IF;
           END_FOR;
           #System.CurrentOrder := 0;
       END_IF;
       IF #Canceling AND NOT (#VTD.Running OR #Extrator_Conveyor.Running OR #Cnv_Buffer_1.Running OR #Cnv_Buffer_2.Running OR #Cnv_Buffer_3.Running) THEN
           #Canceling := FALSE;
           #VTD_CurrentOrder := #Pallet_InOut_CurrentOrder:= #Shuttle_InOut_CurrentOrder := 0;
       END_IF;
   END_REGION

   REGION Resume Orders
       #ResumeRTrig(CLK := #System.ResumeOrders);
       IF #ResumeRTrig.Q THEN
           #System.ResumeOrders := FALSE;
           #System.CurrentOrder := #MaxRunningOrderNo;
           IF NOT #System.Error THEN
               #System.Paused := FALSE;
               FOR #i := 1 TO UDINT_TO_DINT(#MaxRunningOrderNo) DO
                   IF #System.OrderTable[#i].Status = '' THEN
                       EXIT;
                   ELSIF #System.OrderTable[#i].Status = #PAUSED_STATUS
                       OR #System.OrderTable[#i].Status = #ERROR_STATUS
                   THEN
                       #System.OrderTable[#i].Status := #QUEUED_STATUS;
                   END_IF;
               END_FOR;
           END_IF;

       END_IF;
   END_REGION

   REGION Order Handler
       IF #System.Running AND NOT #System.Error
           AND (#System.OrderTable[#System.CurrentOrder].Status = #COMPLETED_STATUS
           OR #System.OrderTable[#System.CurrentOrder].Status = #ERROR_STATUS
           OR #System.OrderTable[#System.CurrentOrder].Status = #ERROR_CANCELED_STATUS
           OR #System.OrderTable[#System.CurrentOrder].Sequence = 0)
       THEN
           IF #System.CurrentOrder > 0 THEN
               #System.CurrentOrder -= 1;
           ELSE
               #System.CurrentOrder := 0;
           END_IF;
       END_IF;
   END_REGION

   REGION Watchdogs
       //Watchdog Timers

       #VTD_WatchdogTimer(IN := #VTD_WatchdogStart,
                          PT := UDINT_TO_TIME(#Watchdog.VTD * 60000),
                          Q => #System.Watchdog_TimeOut.VTD);
       #Pallet_InOut_WatchdogTimer(IN := #Pallet_InOut_WatchdogStart,
                                   PT := UDINT_TO_TIME(#Watchdog.Pallet_INOut * 60000),
                                   Q => #System.Watchdog_TimeOut.Pallet_InOut);
       #Shuttle_InOut_WatchdogTimer(IN := #Shuttle_InOut_WatchdogStart,
                                    PT := UDINT_TO_TIME(#Watchdog.Shuttle_INOut * 60000),
                                    Q => #System.Watchdog_TimeOut.Shuttle_InOut);

       //Reset  Watchdog Timers
       IF #System.Error OR #CancelRTrig.Q OR #PauseRTrig.Q OR "Reset_All" THEN

           #VTD_WatchdogStart := FALSE;
           #Pallet_InOut_WatchdogStart := FALSE;
           #Shuttle_InOut_WatchdogStart := FALSE;

       END_IF;
   END_REGION

   REGION Reset Next Order Number
       IF #System.NextOrder > 1
           AND #CurrentDTL.HOUR = 0
           AND #CurrentDTL.MINUTE = 0
           AND #CurrentDTL.SECOND = 0
       THEN
           #System.NextOrder := 1;
       END_IF;

   END_REGION

   REGION #System Mode and State
       #System.Selected := #System_Selected; // System selected
       #System.Ready := NOT #System.Error AND #System.Selected;
       #System.Auto_Man := #AutoMan_Switch;
       #System.Running :=  #VTD.Running OR #Extrator_Conveyor.Running OR #Cnv_Buffer_1.Running OR #Cnv_Buffer_2.Running OR #Cnv_Buffer_3.Running;

       #System.Error := #VTD.Error OR #Extrator_Conveyor.Error OR #Cnv_Buffer_1.Error OR #Cnv_Buffer_2.Error OR #Cnv_Buffer_3.Error;
       #System.IDLE := NOT #System.Running AND NOT #System.Paused AND NOT #System.Error;
       IF #System.Running THEN
           #System.State := 1;
       ELSIF #System.Paused AND NOT #System.Error THEN
           #System.State := 2;
       ELSIF #System.Error THEN
           #System.State := 3;
       ELSE
           #System.State := 0;
       END_IF;
   END_REGION
END_FUNCTION_BLOCK

FUNCTION "FC_CLOCK" : DTL   // FC55, LAD
{ S7_Optimized_Access := 'TRUE' }
VERSION : 0.1
// stored: AutoNumber true, IsIECCheckEnabled false, SetENOAutomatically false, UDAEnableTagReadback false
   VAR_OUTPUT
      CurrentTime : String;
   END_VAR
   VAR_TEMP
      CurrentDTL : DTL;
      RetVal : Int;
      TempString : String;
      strYear : String;
      strMonth : String;
      strDay : String;
      strHour : String;
      strMinute : String;
      strSeconds : String;
   END_VAR
   VAR_TEMP   // added for the SCL form of the ladder/FBD networks
      _w1 : Bool;
      _w2 : Bool;
      _w3 : Bool;
      _w4 : Bool;
      _w5 : Bool;
   END_VAR
BEGIN

REGION Network 1: Read Current Local Time
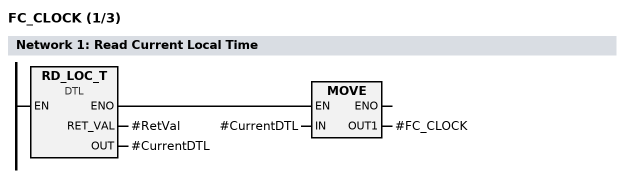
   RUNG wire#powerrail
      { S7_Templates := "date_type := DTL" } RD_LOC_T(RET_VAL => #RetVal, OUT => #CurrentDTL)
      Move(in := #CurrentDTL, out1 => #FC_CLOCK)
   END_RUNG
   // the same network as SCL:
   #RetVal := RD_LOC_T(OUT => #CurrentDTL, ENO => #_w1);
   IF #_w1 THEN #FC_CLOCK := #CurrentDTL; END_IF;
END_REGION

REGION Network 2: Converstion all data to string
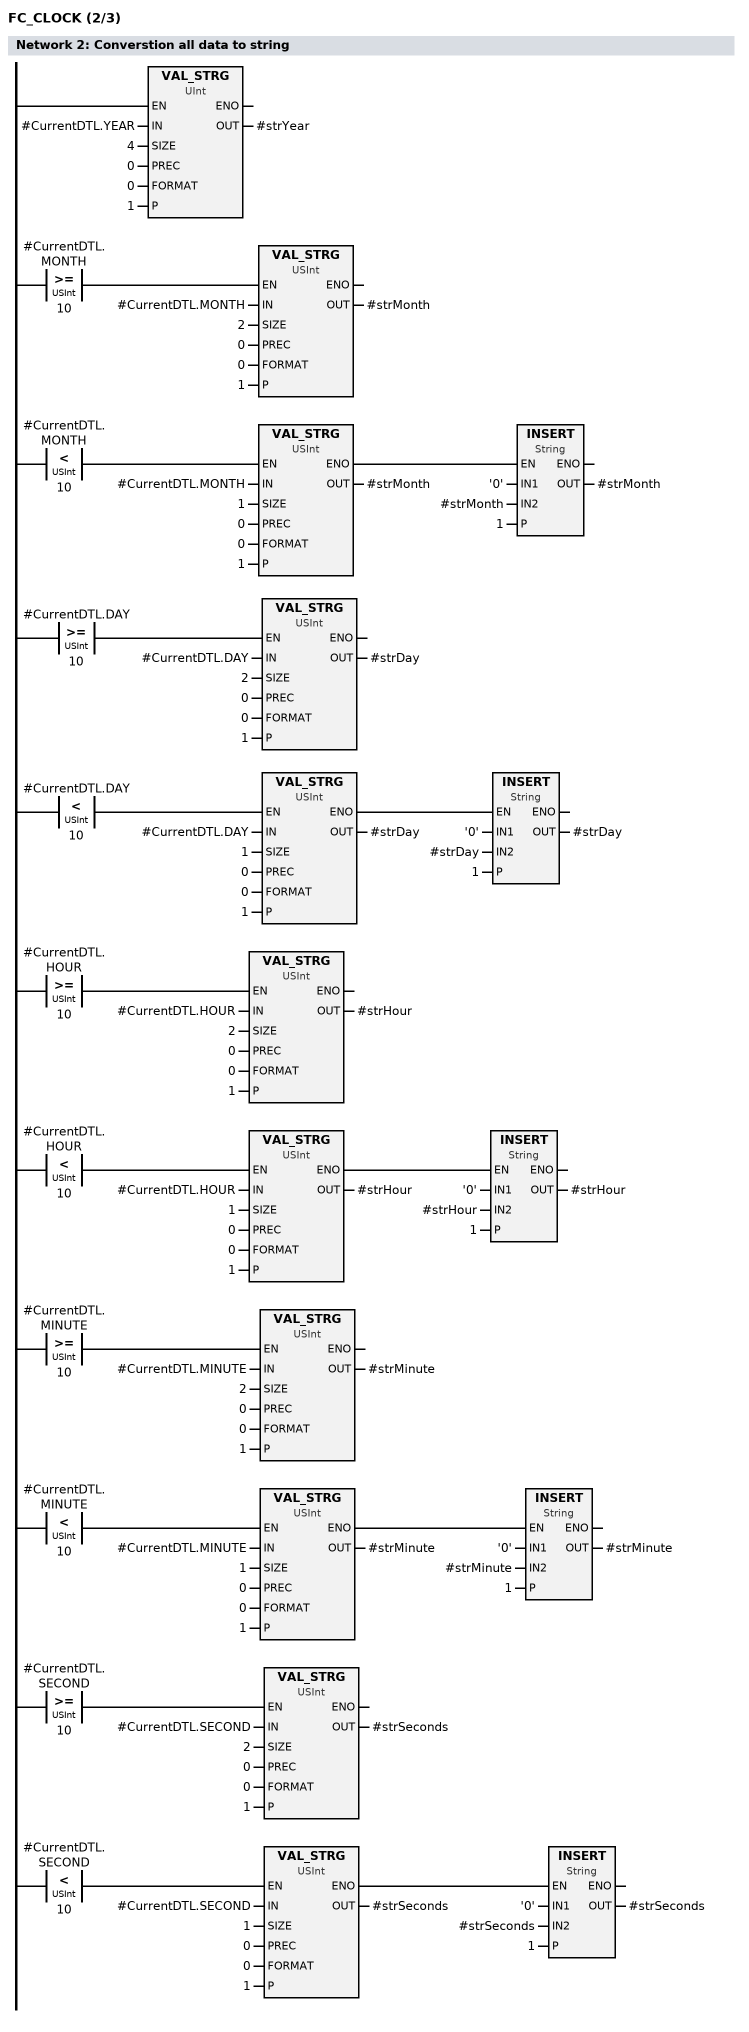
   RUNG wire#powerrail
      { S7_Templates := "[value_type := UInt, str_type := String]" } VAL_STRG(IN := #CurrentDTL.YEAR, SIZE := 4, PREC := 0, FORMAT := 0, P := 1, OUT => #strYear)
   END_RUNG
   RUNG wire#powerrail
      { S7_Templates := "SrcType := USInt" } GE_Contact(in1 := #CurrentDTL.MONTH, in2 := 10)
      { S7_Templates := "[value_type := USInt, str_type := String]" } VAL_STRG(IN := #CurrentDTL.MONTH, SIZE := 2, PREC := 0, FORMAT := 0, P := 1, OUT => #strMonth)
   END_RUNG
   RUNG wire#powerrail
      { S7_Templates := "SrcType := USInt" } LT_Contact(in1 := #CurrentDTL.MONTH, in2 := 10)
      { S7_Templates := "[value_type := USInt, str_type := String]" } VAL_STRG(IN := #CurrentDTL.MONTH, SIZE := 1, PREC := 0, FORMAT := 0, P := 1, OUT => #strMonth)
      { S7_Templates := "str_type := String" } INSERT(IN1 := '0', IN2 := #strMonth, P := 1, OUT => #strMonth)
   END_RUNG
   RUNG wire#powerrail
      { S7_Templates := "SrcType := USInt" } GE_Contact(in1 := #CurrentDTL.DAY, in2 := 10)
      { S7_Templates := "[value_type := USInt, str_type := String]" } VAL_STRG(IN := #CurrentDTL.DAY, SIZE := 2, PREC := 0, FORMAT := 0, P := 1, OUT => #strDay)
   END_RUNG
   RUNG wire#powerrail
      { S7_Templates := "SrcType := USInt" } LT_Contact(in1 := #CurrentDTL.DAY, in2 := 10)
      { S7_Templates := "[value_type := USInt, str_type := String]" } VAL_STRG(IN := #CurrentDTL.DAY, SIZE := 1, PREC := 0, FORMAT := 0, P := 1, OUT => #strDay)
      { S7_Templates := "str_type := String" } INSERT(IN1 := '0', IN2 := #strDay, P := 1, OUT => #strDay)
   END_RUNG
   RUNG wire#powerrail
      { S7_Templates := "SrcType := USInt" } GE_Contact(in1 := #CurrentDTL.HOUR, in2 := 10)
      { S7_Templates := "[value_type := USInt, str_type := String]" } VAL_STRG(IN := #CurrentDTL.HOUR, SIZE := 2, PREC := 0, FORMAT := 0, P := 1, OUT => #strHour)
   END_RUNG
   RUNG wire#powerrail
      { S7_Templates := "SrcType := USInt" } LT_Contact(in1 := #CurrentDTL.HOUR, in2 := 10)
      { S7_Templates := "[value_type := USInt, str_type := String]" } VAL_STRG(IN := #CurrentDTL.HOUR, SIZE := 1, PREC := 0, FORMAT := 0, P := 1, OUT => #strHour)
      { S7_Templates := "str_type := String" } INSERT(IN1 := '0', IN2 := #strHour, P := 1, OUT => #strHour)
   END_RUNG
   RUNG wire#powerrail
      { S7_Templates := "SrcType := USInt" } GE_Contact(in1 := #CurrentDTL.MINUTE, in2 := 10)
      { S7_Templates := "[value_type := USInt, str_type := String]" } VAL_STRG(IN := #CurrentDTL.MINUTE, SIZE := 2, PREC := 0, FORMAT := 0, P := 1, OUT => #strMinute)
   END_RUNG
   RUNG wire#powerrail
      { S7_Templates := "SrcType := USInt" } LT_Contact(in1 := #CurrentDTL.MINUTE, in2 := 10)
      { S7_Templates := "[value_type := USInt, str_type := String]" } VAL_STRG(IN := #CurrentDTL.MINUTE, SIZE := 1, PREC := 0, FORMAT := 0, P := 1, OUT => #strMinute)
      { S7_Templates := "str_type := String" } INSERT(IN1 := '0', IN2 := #strMinute, P := 1, OUT => #strMinute)
   END_RUNG
   RUNG wire#powerrail
      { S7_Templates := "SrcType := USInt" } GE_Contact(in1 := #CurrentDTL.SECOND, in2 := 10)
      { S7_Templates := "[value_type := USInt, str_type := String]" } VAL_STRG(IN := #CurrentDTL.SECOND, SIZE := 2, PREC := 0, FORMAT := 0, P := 1, OUT => #strSeconds)
   END_RUNG
   RUNG wire#powerrail
      { S7_Templates := "SrcType := USInt" } LT_Contact(in1 := #CurrentDTL.SECOND, in2 := 10)
      { S7_Templates := "[value_type := USInt, str_type := String]" } VAL_STRG(IN := #CurrentDTL.SECOND, SIZE := 1, PREC := 0, FORMAT := 0, P := 1, OUT => #strSeconds)
      { S7_Templates := "str_type := String" } INSERT(IN1 := '0', IN2 := #strSeconds, P := 1, OUT => #strSeconds)
   END_RUNG
   // the same network as SCL:
   VAL_STRG(IN := #CurrentDTL.YEAR, SIZE := 4, PREC := 0, FORMAT := 0, P := 1, OUT => #strYear);
   IF #CurrentDTL.MONTH >= 10 THEN
       VAL_STRG(IN := #CurrentDTL.MONTH, SIZE := 2, PREC := 0, FORMAT := 0, P := 1, OUT => #strMonth);
   END_IF;
   VAL_STRG(EN := #CurrentDTL.MONTH < 10,
            IN := #CurrentDTL.MONTH,
            SIZE := 1,
            PREC := 0,
            FORMAT := 0,
            P := 1,
            OUT => #strMonth,
            ENO => #_w1);
   IF #_w1 THEN INSERT(IN1 := '0', IN2 := #strMonth, P := 1, OUT => #strMonth); END_IF;
   IF #CurrentDTL.DAY >= 10 THEN
       VAL_STRG(IN := #CurrentDTL.DAY, SIZE := 2, PREC := 0, FORMAT := 0, P := 1, OUT => #strDay);
   END_IF;
   VAL_STRG(EN := #CurrentDTL.DAY < 10,
            IN := #CurrentDTL.DAY,
            SIZE := 1,
            PREC := 0,
            FORMAT := 0,
            P := 1,
            OUT => #strDay,
            ENO => #_w2);
   IF #_w2 THEN INSERT(IN1 := '0', IN2 := #strDay, P := 1, OUT => #strDay); END_IF;
   IF #CurrentDTL.HOUR >= 10 THEN
       VAL_STRG(IN := #CurrentDTL.HOUR, SIZE := 2, PREC := 0, FORMAT := 0, P := 1, OUT => #strHour);
   END_IF;
   VAL_STRG(EN := #CurrentDTL.HOUR < 10,
            IN := #CurrentDTL.HOUR,
            SIZE := 1,
            PREC := 0,
            FORMAT := 0,
            P := 1,
            OUT => #strHour,
            ENO => #_w3);
   IF #_w3 THEN INSERT(IN1 := '0', IN2 := #strHour, P := 1, OUT => #strHour); END_IF;
   IF #CurrentDTL.MINUTE >= 10 THEN
       VAL_STRG(IN := #CurrentDTL.MINUTE, SIZE := 2, PREC := 0, FORMAT := 0, P := 1, OUT => #strMinute);
   END_IF;
   VAL_STRG(EN := #CurrentDTL.MINUTE < 10,
            IN := #CurrentDTL.MINUTE,
            SIZE := 1,
            PREC := 0,
            FORMAT := 0,
            P := 1,
            OUT => #strMinute,
            ENO => #_w4);
   IF #_w4 THEN INSERT(IN1 := '0', IN2 := #strMinute, P := 1, OUT => #strMinute); END_IF;
   IF #CurrentDTL.SECOND >= 10 THEN
       VAL_STRG(IN := #CurrentDTL.SECOND, SIZE := 2, PREC := 0, FORMAT := 0, P := 1, OUT => #strSeconds);
   END_IF;
   VAL_STRG(EN := #CurrentDTL.SECOND < 10,
            IN := #CurrentDTL.SECOND,
            SIZE := 1,
            PREC := 0,
            FORMAT := 0,
            P := 1,
            OUT => #strSeconds,
            ENO => #_w5);
   IF #_w5 THEN INSERT(IN1 := '0', IN2 := #strSeconds, P := 1, OUT => #strSeconds); END_IF;
END_REGION

REGION Network 3: Current Time String
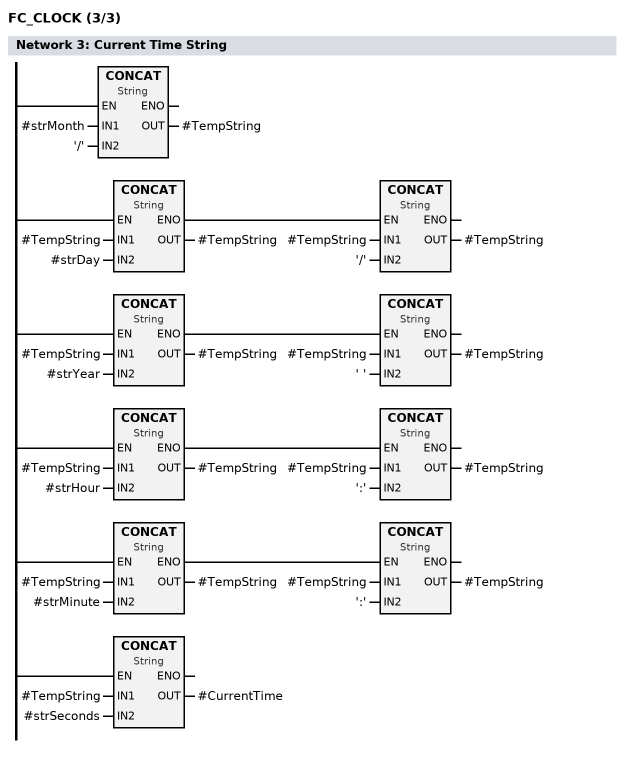
   RUNG wire#powerrail
      { S7_Templates := "[card := 2, str_type := String]" } CONCAT(IN1 := #strMonth, IN2 := '/', OUT => #TempString)
   END_RUNG
   RUNG wire#powerrail
      { S7_Templates := "[card := 2, str_type := String]" } CONCAT(IN1 := #TempString, IN2 := #strDay, OUT => #TempString)
      { S7_Templates := "[card := 2, str_type := String]" } CONCAT(IN1 := #TempString, IN2 := '/', OUT => #TempString)
   END_RUNG
   RUNG wire#powerrail
      { S7_Templates := "[card := 2, str_type := String]" } CONCAT(IN1 := #TempString, IN2 := #strYear, OUT => #TempString)
      { S7_Templates := "[card := 2, str_type := String]" } CONCAT(IN1 := #TempString, IN2 := ' ', OUT => #TempString)
   END_RUNG
   RUNG wire#powerrail
      { S7_Templates := "[card := 2, str_type := String]" } CONCAT(IN1 := #TempString, IN2 := #strHour, OUT => #TempString)
      { S7_Templates := "[card := 2, str_type := String]" } CONCAT(IN1 := #TempString, IN2 := ':', OUT => #TempString)
   END_RUNG
   RUNG wire#powerrail
      { S7_Templates := "[card := 2, str_type := String]" } CONCAT(IN1 := #TempString, IN2 := #strMinute, OUT => #TempString)
      { S7_Templates := "[card := 2, str_type := String]" } CONCAT(IN1 := #TempString, IN2 := ':', OUT => #TempString)
   END_RUNG
   RUNG wire#powerrail
      { S7_Templates := "[card := 2, str_type := String]" } CONCAT(IN1 := #TempString, IN2 := #strSeconds, OUT => #CurrentTime)
   END_RUNG
   // the same network as SCL:
   CONCAT(IN1 := #strMonth, IN2 := '/', OUT => #TempString);
   CONCAT(IN1 := #TempString, IN2 := #strDay, OUT => #TempString, ENO => #_w1);
   IF #_w1 THEN CONCAT(IN1 := #TempString, IN2 := '/', OUT => #TempString); END_IF;
   CONCAT(IN1 := #TempString, IN2 := #strYear, OUT => #TempString, ENO => #_w2);
   IF #_w2 THEN CONCAT(IN1 := #TempString, IN2 := ' ', OUT => #TempString); END_IF;
   CONCAT(IN1 := #TempString, IN2 := #strHour, OUT => #TempString, ENO => #_w3);
   IF #_w3 THEN CONCAT(IN1 := #TempString, IN2 := ':', OUT => #TempString); END_IF;
   CONCAT(IN1 := #TempString, IN2 := #strMinute, OUT => #TempString, ENO => #_w4);
   IF #_w4 THEN CONCAT(IN1 := #TempString, IN2 := ':', OUT => #TempString); END_IF;
   CONCAT(IN1 := #TempString, IN2 := #strSeconds, OUT => #CurrentTime);
END_REGION
END_FUNCTION

FUNCTION_BLOCK "FB_HeartBeat"   // FB25, SCL
{ S7_Optimized_Access := 'TRUE' }
VERSION : 0.1
// stored: AutoNumber true, IsIECCheckEnabled false, IsRetainMemResEnabled false, MemoryReserve 100, SetENOAutomatically false, UDAEnableTagReadback false
   VAR_INPUT
      PC_HeartBeat : Word;
   END_VAR
   VAR_OUTPUT
      PLC_HeartBeat : Word;
      PC_Disconnected : Bool;
   END_VAR
   VAR
      TimeOut : TON_TIME;
      "Timer" { S7_SetPoint := 'True'} : TON_TIME;
      PC_Heartbeat_old : Word;
      StartTimerBit : Bool := FALSE;
   END_VAR
BEGIN
   #Timer(IN := #StartTimerBit, //
          PT := t#500ms);
   IF NOT #StartTimerBit THEN
       #StartTimerBit := TRUE;
   END_IF;
   #Timer(IN := #StartTimerBit, //
          PT := t#500ms);
   IF #Timer.Q THEN
       #StartTimerBit := FALSE;
       RESET_TIMER(#Timer);
       #PLC_HeartBeat += 1;
   END_IF;
   //Time Out Timer
   #TimeOut(IN := #PC_HeartBeat = #PC_Heartbeat_old,
            PT := t#10s);
   #PC_Heartbeat_old := #PC_HeartBeat;
   #PC_Disconnected := #TimeOut.Q; // if time out set PC_Disconnected
END_FUNCTION_BLOCK

